(* IEC 61131-3 sources: daoli-st-library/DL_Motion (part 6) *)

(* ---- FB_DL_AxisCoggingFf.st ---- *)
(*==============================================================================
 * 组件名称 (Component)  : FB_DL_AxisCoggingFf
 * 所属子库 (Sublibrary) : DL_Motion
 * 当前版本 (Version)    : 1.0.0
 * 兼容性   (Platform)   : CODESYS 3.5+ / TwinCAT 3 / 汇川 InoProShop / 施耐德 Machine Expert
 *                         仅依赖 Standard.library（R_TRIG），零厂商私有库
 * 功能描述 (Function)   : 齿槽转矩前馈（按角度周期查表注入）。
 *                         把机械角等分成 72 个扇区（每扇区 5°），表内每格存该角度位置的补偿量；
 *                         运行时按当前角度取格、乘增益、限幅后以转矩前馈输出（% 额定）。
 *                         **学习与注入分离**（互斥锁存）：
 *                           注入态（bInjectEnable）：只读表 + 输出前馈，绝不改表；
 *                           学习态（bLearnEnable） ：只按"实测转矩指令"缓慢更新表内一格，绝不输出前馈；
 *                           两者同拍为真 → 锁存 eLearnConflict 并**两态全停**（既不改表也不输出），
 *                           避免"边学边补"形成正反馈自激。
 *                         三条固化纪律：
 *                           ① **相位取模防越界**：索引由角度除法取整后对 72 取模，负角再补 72，
 *                              结果恒落 0..71；角度非有限或超 ±1E6 度时当拍不判（防整数转换溢出）；
 *                           ② **注入限幅**：输出钳 ±fFfMaxPct，学习后的表格值同样钳在 ±fTableMaxPct；
 *                           ③ **学习率域闸**：fLearnRate 须在 (0, 1] 内，越域即锁存 eCfgIllegal
 *                              （大于 1 的学习率会使表格发散）。
 *                         验收向量：
 *                           ① 角度 0° → 索引 0；角度 5° → 索引 1；角度 355° → 索引 71
 *                           ② 角度 −5° → 索引 71（负角补模）
 *                           ③ 表[0] = 2.0 %、增益 1.0、限幅 5.0 → 前馈 2.0 %
 *                           ④ bInjectEnable 与 bLearnEnable 同拍为真 → eLearnConflict 锁存，输出 0
 * 接口     (Interface)  : 入 fAngleDeg 反馈机械角、bInjectEnable 注入使能、bLearnEnable 学习使能、
 *                         fTorqueRefPct 实测转矩（学习用观测值）、fFfGain 前馈增益、fFfMaxPct 注入限幅、
 *                         fTableMaxPct 表格值限幅、fLearnRate 学习率、bClear 清表沿、bReset 复位沿；
 *                         出 fFfOutPct 转矩前馈输出、iTableIdx 当前表索引（0..71）、bInjecting 注入中、
 *                         bLearning 学习中、bLearnConflict 学/注冲突锁存、bValid 输出有效、
 *                         eState 相、eCause 成因、bError 故障标志。
 * 边界     (Boundary)   : ① **属主边界（写死）：本件只做"角度周期前馈注入与表学习"，不输出位置/速度指令、
 *                         不参与轴使能与故障处理**——与 `FB_DL_AxisFrictionFf` 的分工：齿槽转矩是角度的
 *                         周期函数，摩擦转矩是速度的函数，两表互不替代（R47 边界声明）；
 *                         ② **状态枚举禁定义**：本件不引用任何轴状态枚举（R277），只消费角度引脚；
 *                         ③ **索引边界**：72 格字面量上界（R104），取模后恒在域内，另设显式钳位二次闸；
 *                         ④ **非有限闸**：角度/观测转矩非有限 → 当拍不判、不宣称（不锁存）；
 *                         ⑤ **锁存解除式**：bLearnConflict 与 eFault 仅由 bReset 上升沿解除（R228B），
 *                         bReset 为外部引脚、恒可达；
 *                         ⑥ 零全局耦合、零物理地址。
 * 分工声明 (Scope)      : 本件只管"齿槽转矩前馈"。不接管：摩擦前馈（属 FB_DL_AxisFrictionFf）、
 *                         反向间隙辨识（属 FB_DL_AxisBacklashIdent）、转矩环整定（属驱动侧）。
 * 来源标签 (Source Tag) : 自研线（与 AxisFrictionFf 成族）
 * 码表     (Codes)      : 本件不占用任何全局数字码位（零码位范式 R297）；诊断由 BOOL + ENUM 出口承担。
 * 红线自检 (Redline)    : R1 ✓ 零 GVL/VAR_EXTERNAL ｜ R2 ✓ 零 %I/%Q/%M ｜ R3 ✓ 纯 IEC 61131-3
 *                         R4 ✓ 取模 + 显式钳位 + 双限幅 + 学习率域闸 + 非有限闸 ｜ R5 ✓ 声明逐行同行双语注释
 *                         R6 ✓ ENUM+CASE 含 ELSE 兜底 ｜ R7 ✓ 两 R_TRIG 段 0 无条件刷新（本件无 TON）
 * 修订历史 (Revision)   : 2026-11-19  v1.0.0  R47 首版（批次 4 · 序号 20）
 *==============================================================================*)

TYPE E_DL_AcgState :
(
    eIdle  := 0,    // 待机相（两态皆关，输出 0） / Idle, both modes off, zero output
    eInject:= 10,   // 注入相（只读表输出前馈） / Injecting, table read only
    eLearn := 20,   // 学习相（只更新表，无输出） / Learning, table update only
    eFault := 90    // 故障相（等复位） / Fault, awaiting reset
);
END_TYPE

TYPE E_DL_AcgCause :
(
    eNone         := 0,   // 无异常 / No anomaly
    eCfgIllegal   := 1,   // 组态非法（学习率/限幅越域） / Illegal configuration
    eLearnConflict:= 2,   // 学习与注入同拍（锁存，两态全停） / Learn and inject together, latched
    eAngleBad     := 3,   // 角度非有限或超域（当拍不判） / Angle invalid, skipped this scan
    ePhaseBad     := 4    // 非法相位兜底 / Illegal phase fallback
);
END_TYPE

FUNCTION_BLOCK FB_DL_AxisCoggingFf
VAR_INPUT
    fAngleDeg    : LREAL := 0.0;      // 反馈机械角（可正可负） [°] / Feedback mechanical angle [°]
    bInjectEnable: BOOL := FALSE;     // 注入使能（只读表） [-] / Injection enable, table read only
    bLearnEnable : BOOL := FALSE;     // 学习使能（只改表） [-] / Learning enable, table write only
    fTorqueRefPct: LREAL := 0.0;      // 实测转矩（学习观测值） [% 额定] / Measured torque for learning [% rated]
    fFfGain      : LREAL := 1.0;      // 前馈增益，域 ≥ 0 [-] / Feed-forward gain, >= 0
    fFfMaxPct    : LREAL := 20.0;     // 注入限幅，域 > 0 [% 额定] / Injection clamp, > 0
    fTableMaxPct : LREAL := 30.0;     // 表格值限幅，域 > 0 [% 额定] / Table-value clamp, > 0
    fLearnRate   : LREAL := 0.01;     // 学习率，域 (0, 1] [-] / Learning rate, within (0, 1]
    bClear       : BOOL := FALSE;     // 清表沿（表格全置 0） [-] / Table-clear edge
    bReset       : BOOL := FALSE;     // 故障复位沿 [-] / Fault reset edge
END_VAR
VAR_OUTPUT
    fFfOutPct    : LREAL := 0.0;                          // 转矩前馈输出（已限幅） [% 额定] / Feed-forward output, clamped
    iTableIdx    : INT := 0;                              // 当前表索引（0..71） [-] / Present table index
    bInjecting   : BOOL := FALSE;                         // 注入中 [-] / Injecting
    bLearning    : BOOL := FALSE;                         // 学习中 [-] / Learning
    bLearnConflict : BOOL := FALSE;                       // 学/注冲突锁存（等复位） [-] / Learn-inject conflict, latched
    bValid       : BOOL := FALSE;                         // 输出有效（角度有效且注入态） [-] / Output valid
    eState       : E_DL_AcgState := E_DL_AcgState.eIdle;  // 相出口 [-] / Phase outlet
    eCause       : E_DL_AcgCause := E_DL_AcgCause.eNone;  // 成因出口（R190 归因唯一） [-] / Cause outlet
    bError       : BOOL := FALSE;                         // 故障标志（仅故障级成因） [-] / Error flag, fault level only
END_VAR
VAR
    _eState   : E_DL_AcgState := E_DL_AcgState.eIdle;    // 内部相（CASE 唯一写入目标） / Internal phase
    _eCause   : E_DL_AcgCause := E_DL_AcgCause.eNone;    // 成因锁存量 / Latched cause
    _bFault   : BOOL := FALSE;                           // 故障锁存位 / Latched fault bit
    _bConf    : BOOL := FALSE;                           // 学/注冲突锁存位 / Latched conflict bit
    _iIdx     : INT := 0;                                // 归一后的表索引（0..71） [-] / Normalised table index
    _iRaw     : INT := 0;                                // 取模前的索引 [-] / Index before normalisation
    _fOut     : LREAL := 0.0;                            // 输出工作值 [% 额定] / Output working value
    _fCell    : LREAL := 0.0;                            // 当格补偿量 [% 额定] / Cell compensation value
    _bAngOk   : BOOL := FALSE;                           // 角度有效性结论 / Angle validity result
    _bCfgBad  : BOOL := FALSE;                           // 组态非法当拍量 / Illegal configuration this scan
    _i        : INT := 0;                                // 清表循环下标 / Clear-loop index
    rtClear   : R_TRIG;                                  // 清表沿实例，段 0 无条件调用 / Clear edge instance
    rtReset   : R_TRIG;                                  // 复位沿实例，段 0 无条件调用 / Reset edge instance
    afTable   : ARRAY[0..71] OF LREAL;                   // 齿槽补偿表（72 格 = 5°/格，字面量上界） [% 额定] / Cogging table
END_VAR
VAR CONSTANT
    DL_ACG_NBINS   : INT := 72;          // 表格数（与数组字面量上界同源） [格] / Table bin count
    DL_ACG_BIN_DEG : LREAL := 5.0;       // 每格角度宽（360/72） [°] / Bin width in degrees
    DL_ACG_ANG_MAX : LREAL := 1000000.0; // 角度绝对值上限（防实数转整数溢出） [°] / Angle magnitude limit
    DL_ACG_EPS     : LREAL := 1.0E-12;   // 浮点判等容差 [-] / Equality tolerance
END_VAR

(* —— 段 0：组态闸 + 两沿无条件周期刷新（R228A；本件无 TON） —— *)
_bCfgBad := (fLearnRate <= 0.0) OR (fLearnRate > 1.0)                 // 学习率须在 (0, 1] / Learning rate within (0, 1]
         OR (fFfMaxPct <= 0.0) OR (fTableMaxPct <= 0.0)               // 两限幅须为正 / Both clamps positive
         OR (fFfGain < 0.0);                                          // 增益须非负 / Gain non-negative
rtClear(CLK := bClear);                                               // 清表沿 / Clear edge
rtReset(CLK := bReset);                                               // 复位沿 / Reset edge

(* —— 段 1：单拍/输出量预置（锁存量 _eCause/_bFault/_bConf/_iIdx 不入清单，R107） —— *)
fFfOutPct  := 0.0;                                                    // 前馈输出预置 / Feed-forward preset
bInjecting := FALSE;                                                  // 注入中预置 / Injecting preset
bLearning  := FALSE;                                                  // 学习中预置 / Learning preset
bValid     := FALSE;                                                  // 有效位预置 / Validity preset
bError     := FALSE;                                                  // 故障标志预清（R45 配对） / Error preset
_fOut      := 0.0;                                                    // 输出工作值预置 / Output working preset

(* —— 段 2：组态闸（非法即锁存） —— *)
IF _bCfgBad THEN
    _eCause := E_DL_AcgCause.eCfgIllegal;                             // 归因：组态非法 / Cause: illegal configuration
    _bFault := TRUE;                                                  // 锁存 / Latch
    _eState := E_DL_AcgState.eFault;                                  // 入故障相 / Enter fault phase
END_IF

(* —— 段 3：学/注冲突闸（同拍为真即锁存，两态全停） —— *)
IF bInjectEnable AND bLearnEnable THEN
    _bConf  := TRUE;                                                  // 冲突锁存 / Latch the conflict
    _bFault := TRUE;                                                  // 故障锁存 / Latch the fault
    _eCause := E_DL_AcgCause.eLearnConflict;                          // 归因：学/注冲突 / Cause: learn-inject conflict
    _eState := E_DL_AcgState.eFault;                                  // 入故障相 / Enter fault phase
END_IF

(* —— 段 4：迁出链与清表链（两条显式写出） —— *)
IF rtReset.Q THEN
    _bFault := FALSE;                                                 // 清故障锁存 / Clear fault latch
    _bConf  := FALSE;                                                 // 清冲突锁存 / Clear the conflict latch
    _eCause := E_DL_AcgCause.eNone;                                   // 清成因 / Clear cause
    _eState := E_DL_AcgState.eIdle;                                   // 回待机相 / Back to idle
END_IF
IF rtClear.Q THEN
    FOR _i := 0 TO 71 DO
        afTable[_i] := 0.0;                                           // 逐格清零（循环上界恒定） / Clear every bin
    END_FOR
END_IF

(* —— 段 5：索引归一（角度有限性 → 取整 → 取模 → 负角补模 → 显式钳位） —— *)
_bAngOk := NOT ((fAngleDeg <> fAngleDeg) OR ((fAngleDeg - fAngleDeg) <> (fAngleDeg - fAngleDeg)))
        AND (ABS(fAngleDeg) <= DL_ACG_ANG_MAX);                       // 有限且未超防溢出上限 / Finite and below the guard limit
IF _bAngOk THEN
    _iRaw := LREAL_TO_INT(TRUNC(fAngleDeg / DL_ACG_BIN_DEG));         // 取整到格号（截断向 0） / Truncate to a bin number
    _iIdx := _iRaw MOD DL_ACG_NBINS;                                  // 对格数取模 / Modulo the bin count
    IF _iIdx < 0 THEN
        _iIdx := _iIdx + DL_ACG_NBINS;                                // 负角补模（−5° → 71） / Negative angle wrapped
    END_IF
    IF _iIdx < 0 THEN
        _iIdx := 0;                                                   // 二次下钳（结构性冗余） / Second lower clamp
    ELSIF _iIdx > (DL_ACG_NBINS - 1) THEN
        _iIdx := DL_ACG_NBINS - 1;                                    // 二次上钳（结构性冗余） / Second upper clamp
    END_IF
    iTableIdx := _iIdx;                                               // 索引出口 / Index outlet
ELSE
    _eCause := E_DL_AcgCause.eAngleBad;                               // 归因：角度无效（当拍不判） / Cause: invalid angle
END_IF

(* —— 段 6：相迁移（注入 / 学习互斥；故障由段 4 迁出） —— *)
CASE _eState OF

E_DL_AcgState.eIdle:
    IF bInjectEnable AND (NOT bLearnEnable) THEN
        _eState := E_DL_AcgState.eInject;                              // 进注入相 / Enter injecting
    ELSIF bLearnEnable AND (NOT bInjectEnable) THEN
        _eState := E_DL_AcgState.eLearn;                               // 进学习相 / Enter learning
    END_IF

E_DL_AcgState.eInject:
    IF bLearnEnable THEN
        _eState := E_DL_AcgState.eIdle;                                // 学习被使能：先退注入（互斥由段 3 判冲突） / Leave injecting
    ELSIF NOT bInjectEnable THEN
        _eState := E_DL_AcgState.eIdle;                                // 失能：回待机 / Disabled, back to idle
    END_IF

E_DL_AcgState.eLearn:
    IF bInjectEnable THEN
        _eState := E_DL_AcgState.eIdle;                                // 注入被使能：先退学习 / Leave learning
    ELSIF NOT bLearnEnable THEN
        _eState := E_DL_AcgState.eIdle;                                // 失能：回待机 / Disabled, back to idle
    END_IF

E_DL_AcgState.eFault:
    ;                                                                  // 故障相：由段 4 复位沿迁出 / Exit via the reset edge

ELSE
    _eCause := E_DL_AcgCause.ePhaseBad;                                // 归因：非法相位 / Cause: illegal phase
    _bFault := TRUE;                                                   // 锁存 / Latch
    _eState := E_DL_AcgState.eFault;                                   // 强拉故障相 / Force fault phase

END_CASE

(* —— 段 7：注入（只读表；增益与限幅） —— *)
IF (_eState = E_DL_AcgState.eInject) AND _bAngOk THEN
    _fCell := afTable[_iIdx];                                           // 读当格补偿量 / Read the cell value
    _fOut  := _fCell * fFfGain;                                         // 乘增益 / Apply the gain
    IF _fOut > fFfMaxPct THEN
        _fOut := fFfMaxPct;                                             // 上限钳位 / Clamp high
    ELSIF _fOut < (0.0 - fFfMaxPct) THEN
        _fOut := 0.0 - fFfMaxPct;                                       // 下限钳位 / Clamp low
    END_IF
    bInjecting := TRUE;                                                 // 注入中 / Injecting
    bValid     := TRUE;                                                 // 输出有效 / Output valid
END_IF

(* —— 段 8：学习（只改表；观测转矩有限才更新；表值双限幅） —— *)
IF (_eState = E_DL_AcgState.eLearn) AND _bAngOk THEN
    IF NOT ((fTorqueRefPct <> fTorqueRefPct) OR ((fTorqueRefPct - fTorqueRefPct) <> (fTorqueRefPct - fTorqueRefPct))) THEN
        afTable[_iIdx] := afTable[_iIdx] + (fLearnRate * fTorqueRefPct);   // 梯度式更新（学习率已过域闸） / Gradient-style update
        IF afTable[_iIdx] > fTableMaxPct THEN
            afTable[_iIdx] := fTableMaxPct;                             // 表格上限钳位 / Table clamp high
        ELSIF afTable[_iIdx] < (0.0 - fTableMaxPct) THEN
            afTable[_iIdx] := 0.0 - fTableMaxPct;                       // 表格下限钳位 / Table clamp low
        END_IF
        bLearning := TRUE;                                              // 学习中 / Learning
    END_IF
END_IF

(* —— 段 9：出口单点映射（名实双出口，R191） —— *)
fFfOutPct      := _fOut;                                                // 前馈输出出口 / Feed-forward outlet
bLearnConflict := _bConf;                                               // 冲突锁存出口 / Conflict outlet
eState         := _eState;                                              // 相出口 / Phase outlet
eCause         := _eCause;                                              // 成因出口 / Cause outlet
bError         := _bFault;                                              // 故障标志 / Error flag

END_FUNCTION_BLOCK

(* ---- FB_DL_AxisDroopComp.st ---- *)
(*==============================================================================
 * 组件名称 (Component)  : FB_DL_AxisDroopComp
 * 所属子库 (Sublibrary) : DL_Motion
 * 当前版本 (Version)    : 1.0.0
 * 兼容性   (Platform)   : CODESYS 3.5 / TwinCAT 3 / 汇川 InoProShop / Machine Expert
 *                         仅依赖 Standard.library（R_TRIG），零厂商方言
 * 功能描述 (Function)   : 轴跟随误差前馈补偿：按速度段从补偿表取增益，折算位置前置量
 *                         fCompOut [mm] = 速度段增益 [mm per mm/s] × 速度给定 [mm/s]，
 *                         并钳在 ±fCompMax；用于抵消伺服刚度不足造成的跟随下垂。
 * 分工互引 (Boundary)   : FB_DL_AxisFollowErrGuard 是**保护件**（跟随误差超限即停），
 *                         本件是**补偿件**（前置量注入位置环，不产生任何停止动作）；
 *                         两者互不替代，禁把保护判据写进本件。
 *                         FB_DL_AxisFrictionFf 补偿摩擦力方向项，本件只补偿速度相关下垂。
 * 边界与语义披露 (Boundary disclosure) :
 *   1) 补偿表 8 段定长（DL_AC_SEG），段边界按 |fVelCmd| 等分 fVelSegMax，
 *      符号由速度给定方向携带（段内取绝对值查表，输出乘回方向），故负速也有补偿。
 *   2) 组态域闸（R151 全枚举）：fVelSegMax <= 0、fCompMax < 0、表内任一元素非有限或
 *      为负（负增益会让补偿反向加剧下垂）均判组态非法，锁存至复位沿 + 组态改对。
 *   3) 速度给定非有限属运行时信号失效：本拍不输出补偿（fCompOut := 0，安全侧不注入
 *      错误前置量），置信息级码，**不锁存**（不因一扫 NaN 让补偿永久失效）。
 *   4) 输出饱和（|补偿| 被 fCompMax 钳住）为信息级：饱和本身不改变补偿符号。
 * 故障码表 (Error codes) :
 *   16#0004_03F0 [故障级] 组态非法（段宽 / 补偿上限 / 表元素），补偿置 0
 *                 反证：补偿置 0 与「速度恰好为 0」输出组合相同，无码不可区分。
 *   16#0004_03F2 [信息级] 速度给定非有限，本拍不注入补偿（保持 0）
 *                 反证：补偿 0 与「低速段增益为 0」输出相同，需码位区分信号失效。
 *   16#0004_03F3 [信息级] 补偿量被上限钳位（bSaturated 同源可查）
 *                 反证：钳位后补偿与前一段恰好相同，无码不可观测。
 * 码位总账 (Code ledger) : 16#0004_03F0 用 ｜ 16#0004_03F2 / 03F3 用
 * 依赖     (Depends)    : 无 DL_ 内部依赖；Standard.library: R_TRIG
 * 红线自检 (Redline)    : R1 ✓ 零全局变量 ｜ R2 ✓ 零 %I/%Q ｜ R3 ✓ 纯 IEC 61131-3
 *                         R4 ✓ 段索引钳位无越界 / 非有限三判 / 除子由域闸保证 > 0
 *                         R5 ✓ 全变量双语同行注释 ｜ R6 ✓ 三态 ENUM + ELSE 兜底
 *                         R7 ✓ 一沿实例主体最前部无条件刷新
 * 修订历史 (Revision)   : 2026-11-22  v1.0.0  首版入库（R69 构建轮 · 批 3 · N8）
 *============================================================================*)

(*-----------------------------------------------------------------------------
 * 枚举: E_DL_DroopState（归属 DL_Motion，与 FB_DL_AxisDroopComp 同文件）
 *----------------------------------------------------------------------------*)
TYPE E_DL_DroopState :
(
    eOff   := 0,      // 未使能：补偿恒 0 / Disabled, compensation is zero
    eRun   := 10,     // 补偿中：按速度段查表 / Compensating by speed segment
    eFault := 99      // 组态锁存：补偿恒 0 / Config latched, compensation forced to zero
);
END_TYPE

(*==============================================================================
 * 功能块: FB_DL_AxisDroopComp
 * 调用约定: 每个扫描周期无条件调用一次。
 *============================================================================*)
FUNCTION_BLOCK FB_DL_AxisDroopComp
VAR_INPUT
    fVelCmd    : REAL;                          // 速度给定 [mm/s] / velocity setpoint [mm/s]
    afSegGain  : ARRAY[0..7] OF REAL;           // 8 段补偿增益 [mm per mm/s]，必须 >= 0 / per-segment droop gain
    fVelSegMax : REAL := 1000.0;                // 补偿表覆盖的最高速度 [mm/s]，<= 0 组态非法 / table velocity span
    fCompMax   : REAL := 2.0;                   // 补偿量上限 [mm]，< 0 组态非法 / compensation magnitude ceiling [mm]
    bEnable    : BOOL := TRUE;                  // 使能 / enable
    bReset     : BOOL;                          // 上升沿：清组态锁存 / rising edge clears the config latch
END_VAR
VAR_OUTPUT
    fCompOut   : REAL;                          // 位置前置补偿量 [mm]（含速度方向符号）/ position feed-forward [mm]
    nSegIdx    : INT;                           // 命中补偿段号 [段]，0..7 / hit segment index
    bSaturated : BOOL;                          // 补偿量被上限钳位 / compensation clamped at the ceiling
    bVelValid  : BOOL;                          // 本拍速度给定有限 / velocity setpoint finite this scan
    bError     : BOOL;                          // 故障标志（组态锁存）/ fault flag
    uErrorId   : UDINT;                         // 故障码，0 = 无故障 / error code, 0 = none
    eState     : E_DL_DroopState;               // 当前状态（供 HMI 诊断）/ current state
END_VAR
VAR
    fbTrigReset : R_TRIG;                       // 复位沿检测实例 / reset edge detector
    eStateInt   : E_DL_DroopState;              // 主状态机内部当前态 / internal state
    fVelAbs     : REAL;                         // 速度绝对值 [mm/s]（查表用）/ absolute velocity for the lookup
    fSegSpan    : REAL;                         // 单段速度宽度 [mm/s]（除子，域闸保证 > 0）/ segment width, the divisor
    fGainEff    : REAL;                         // 命中段增益 [mm per mm/s] / hit segment gain
    fCompRaw    : REAL;                         // 未钳补偿量 [mm] / unclamped compensation
    nIdx        : INT;                          // 表遍历游标 [段] / table cursor
    bVelBad     : BOOL;                         // 速度给定非有限 / velocity non-finite
    bCfgBad     : BOOL;                         // 本拍组态非法 / config illegal this scan
    bCfgLatch   : BOOL;                         // 组态锁存（复位沿 + 组态改对解除）/ config latch
    bErrorInt   : BOOL;                         // 本拍故障置位累加 / fault set accumulator
    bFirstScan  : BOOL := TRUE;                 // 上电首扫标志 / first-scan flag
END_VAR
VAR CONSTANT
    DL_AC_SEG     : INT := 8;                   // 补偿表段数 [段]，与数组维度一致 / segment count
    DL_AC_FIN_LIM : REAL := 1.0E30;             // REAL 幅值兜底判界 / REAL magnitude bound
    DL_AC_NEG_EPS : REAL := 0.0;                // 增益负值判界（0 为合法端点）/ gain negativity bound, zero is legal
END_VAR

(*------------------------------------------------------------------------------
 * 段 1｜无条件刷新区（红线 R7）：一沿实例位于主体最前部
 *      Unconditional refresh: the edge instance at the very top
 *-----------------------------------------------------------------------------*)
fbTrigReset(CLK := bReset);

(* 段 2｜上电首扫：状态与输出落安全侧 / first-scan init *)
IF bFirstScan THEN
    eStateInt  := E_DL_DroopState.eOff;
    fCompOut   := 0.0;
    bFirstScan := FALSE;
END_IF

(* 段 3｜每拍预清（FB32-1）：单拍标志与派生量 / per-scan preset *)
bErrorInt  := FALSE;
bSaturated := FALSE;

(*------------------------------------------------------------------------------
 * 段 4｜组态域闸（R151 全枚举）：段宽 / 上限 / 表内 8 个元素逐一非有限与负值判
 *      Config gate over the span, the ceiling and every table element
 *      解除路径（R152 自证可达）：复位沿 AND 组态非法条件全部消失
 *-----------------------------------------------------------------------------*)
bCfgBad := (fVelSegMax <= 0.0) OR (fVelSegMax <> fVelSegMax)
           OR (fCompMax < 0.0) OR (fCompMax <> fCompMax);
FOR nIdx := 0 TO (DL_AC_SEG - 1) DO
    IF (afSegGain[nIdx] <> afSegGain[nIdx])
       OR ((afSegGain[nIdx] - afSegGain[nIdx]) <> (afSegGain[nIdx] - afSegGain[nIdx]))
       OR (ABS(afSegGain[nIdx]) >= DL_AC_FIN_LIM)
       OR (afSegGain[nIdx] < DL_AC_NEG_EPS) THEN
        bCfgBad := TRUE;                        // 表元素非法：任一项即整表不可信 / any bad element invalidates the table
    END_IF
END_FOR

IF bCfgBad THEN
    bCfgLatch := TRUE;
END_IF
IF fbTrigReset.Q AND (NOT bCfgBad) THEN
    bCfgLatch := FALSE;                         // 组态锁存解除 / config latch cleared
    uErrorId  := 16#0000_0000;                  // 码位随解除归零 / code cleared with the latch
END_IF
IF bCfgLatch THEN
    uErrorId  := 16#0004_03F0;                  // 故障级：组态非法 / fault: illegal configuration
    bErrorInt := TRUE;                          // R45 配对 / paired with the code
    eStateInt := E_DL_DroopState.eFault;
END_IF

(*------------------------------------------------------------------------------
 * 段 5｜主状态机（红线 R6）：ENUM + CASE + ELSE 兜底
 *-----------------------------------------------------------------------------*)
CASE eStateInt OF

    E_DL_DroopState.eOff:
        IF bEnable AND (NOT bCfgLatch) THEN
            eStateInt := E_DL_DroopState.eRun;
        END_IF

    E_DL_DroopState.eRun:
        IF (NOT bEnable) OR bCfgLatch THEN
            eStateInt := E_DL_DroopState.eOff;
        END_IF

    E_DL_DroopState.eFault:
        IF fbTrigReset.Q AND (NOT bCfgBad) THEN
            bCfgLatch := FALSE;
            uErrorId  := 16#0000_0000;
            eStateInt := E_DL_DroopState.eOff;
        END_IF

    ELSE
        (* 非法状态拦截 / illegal state interception *)
        eStateInt := E_DL_DroopState.eFault;
        uErrorId  := 16#0004_03F0;
        bErrorInt := TRUE;

END_CASE;

(*------------------------------------------------------------------------------
 * 段 6｜速度段查表与补偿折算
 *      Segment lookup and the compensation folding
 *-----------------------------------------------------------------------------*)
bVelBad  := (fVelCmd <> fVelCmd)
            OR ((fVelCmd - fVelCmd) <> (fVelCmd - fVelCmd))
            OR (ABS(fVelCmd) >= DL_AC_FIN_LIM);
bVelValid := (NOT bVelBad) AND (NOT bCfgLatch);
fCompOut  := 0.0;                               // 缺省不注入（安全侧）/ default no injection
nSegIdx   := 0;
fGainEff  := 0.0;

IF bVelValid AND bEnable AND (eStateInt = E_DL_DroopState.eRun) THEN
    IF fVelCmd >= 0.0 THEN
        fVelAbs := fVelCmd;                     // 正方向 [mm/s] / positive direction
    ELSE
        fVelAbs := -fVelCmd;                    // 取绝对值查表（符号在出口乘回）[mm/s] / absolute value for the lookup
    END_IF
    fSegSpan := fVelSegMax / INT_TO_REAL(DL_AC_SEG);                 // 单段宽（除子为常数 8 > 0）[mm/s] / segment width
    IF fVelAbs > fVelSegMax THEN
        fVelAbs := fVelSegMax;                  // 实数域先钳制再转整型（R151 防方向翻转）/ clamp in the real domain before the cast
    END_IF
    nSegIdx  := REAL_TO_INT(fVelAbs / fSegSpan);                     // 段号（除子 > 0 且已钳制）/ segment index after clamping
    IF nSegIdx >= DL_AC_SEG THEN
        nSegIdx := DL_AC_SEG - 1;               // 超表按末段钳位（禁越界访问）/ clamp to the last segment
    ELSIF nSegIdx < 0 THEN
        nSegIdx := 0;                           // 负段号防御，结构性不可达 / negative guard, unreachable
    END_IF
    fGainEff := afSegGain[nSegIdx];             // 命中段增益 [mm per mm/s] / hit gain
    fCompRaw := fGainEff * fVelCmd;             // 未钳补偿（含方向符号）[mm] / raw compensation with direction
    IF fCompRaw > fCompMax THEN
        fCompOut   := fCompMax;                 // 正向饱和 [mm] / saturated high
        bSaturated := TRUE;
        uErrorId   := 16#0004_03F3;             // 信息级：补偿被钳位 / info: compensation clamped
    ELSIF fCompRaw < -fCompMax THEN
        fCompOut   := -fCompMax;                // 负向饱和 [mm] / saturated low
        bSaturated := TRUE;
        uErrorId   := 16#0004_03F3;             // 信息级：补偿被钳位 / info: compensation clamped
    ELSE
        fCompOut   := fCompRaw;                 // 域内直通 [mm] / in-domain pass-through
    END_IF
ELSIF bVelBad THEN
    uErrorId := 16#0004_03F2;                   // 信息级：速度非有限，不注入（不锁存）/ info: non-finite velocity
END_IF

(*------------------------------------------------------------------------------
 * 段 7｜输出单一出口（范式 P-05）
 *      Single output exit
 *-----------------------------------------------------------------------------*)
bError := bErrorInt OR bCfgLatch;
eState := eStateInt;
END_FUNCTION_BLOCK

(* ---- FB_DL_AxisDualFeedbackGuard.st ---- *)
(*==============================================================================
 * 组件名称 (Component)  : FB_DL_AxisDualFeedbackGuard
 * 所属子库 (Sublibrary) : DL_Motion
 * 当前版本 (Version)    : 1.0.0
 * 兼容性   (Platform)   : CODESYS 3.5+ / TwinCAT 3 / 汇川 InoProShop / 施耐德 Machine Expert
 *                         仅依赖 Standard.library（TON / R_TRIG / ABS），零厂商私有库
 * 功能描述 (Function)   : 单轴双反馈交叉校核。把电机侧位置 fPosMotor 与负载侧位置 fPosLoad
 *                         各自乘标定系数换算到同一工程单位后求偏差 fDev，并按幅值与持续时间
 *                         分级：|fDev| 超 fDevWarn → 维护级预警（bWarn）；超 fDevAlarm 且持续
 *                         tDevConfirm → 故障锁存。另做极性装反识别：偏差方向与参考运动方向
 *                         同号、且偏差每拍增量超 fSlopeThr 时归因 ePolarity（区别于打滑——
 *                         打滑时偏差随运动累积但方向与运动一致而增量平稳，装反时增量陡增）。
 * 接口     (Interface)  : 输入 fPosMotor 电机侧位置、fPosLoad 负载侧位置、fScaleMotor / fScaleLoad
 *                         两侧标定系数、fDevWarn 预警阈值、fDevAlarm 故障阈值、tDevConfirm 故障
 *                         确认时间、fSlopeThr 偏差每拍增量阈值、fVelRefMms 参考运动速度（方向
 *                         判据）、bReset 复位；输出 fDev 换算后偏差、bWarn 维护级预警、bGuardOk
 *                         校核通过、eState / eCause / bError / nErrId。
 * 边界     (Boundary)   : ① 组态闸：fScaleMotor / fScaleLoad 的绝对值 <= DL_FLOAT_EPS（防零增益
 *                         静默把偏差算成 0）、fDevWarn <= 0.0、fDevAlarm <= fDevWarn、
 *                         tDevConfirm <= T#0S、fSlopeThr < 0.0 或任一浮点引脚 NaN → 故障锁存；
 *                         ② **本件不定义轴状态枚举、不发运动指令**（轴状态唯一属主 `I_DL_MotionAxis`），
 *                         只读位置与速度参考，只输出校核结论；
 *                         ③ 偏差每拍增量以「每拍工程单位增量」为单位：任务周期固定时它与斜率
 *                         成正比，fSlopeThr 按该口径标定（比值约定见头注释遗留假设）；
 *                         ④ TON 两枚（预警/故障确认）+ R_TRIG 一枚段 0 无条件周期刷新；
 *                         ⑤ 故障相迁出唯一路径 = bReset 上升沿；⑥ 零全局耦合（无 GVL / 无物理地址）。
 * 分工声明 (Scope)      : 与 `FB_DL_GantrySyncAxis`（双**轴**同步偏差）分工 —— 本件是**单轴双反馈**
 *                         （电机侧 vs 负载侧），判「同一根轴的两把尺是否一致」；那件判「两根轴的
 *                         位置是否同步」。二者输入维度不同，禁止互相替代。
 * 遗留假设 (Assumption) : 【R95 三句声明】① 代理值 = 偏差每拍增量（未引入任务周期引脚）；
 *                         ② 覆盖范围 = 任务周期 1 ms ~ 20 ms 的常规运动任务；③ 覆盖不到的区间
 *                         （< 1 ms 的高速插补任务）由调用方负责：此时每拍增量被任务周期压缩，
 *                         fSlopeThr 需由调用方按周期比例放大，否则极性识别灵敏度下降。
 * 解除式   (Release)    : bReset 上升沿 ∧ 组态合法 ∧ |fDev| < fDevWarn（当拍量，R240 范式）。
 *                         自证可满足（终审两式 1）：解除式只含当拍偏差比较与组态闸，两枚 TON
 *                         的 IN 由当拍阈值判据派生，偏差回落即 Q 落假，无恒假因子。
 * 码表     (Codes)      : 16#0004_03B4 故障级：双反馈校核故障总码（组态非法 / 偏差超限确认 /
 *                         极性装反 / 非法相位），锁存至 bReset 上升沿，归因由 eCause 承载；
 *                         16#0004_04B4 信息级：维护级预警（|fDev| 超 fDevWarn 但未达故障）。
 *                         加码反证（R90）：预警相 fDev 仍为小值、bError 为假，若只靠 bWarn 布尔
 *                         位则该退化不进报警台账（HMI 只归档带码事件），故立一码。
 *                         码段说明：0004 段故障子带 03xx / 信息子带 04xx，本件取 03B4 / 04B4
 *                         （源码实扫该两槽为空，续接同子带已用最大值，未回填碎片孔洞）。
 * 开源溯源 (Origin)     : 道莅自研 clean-room（参考双反馈交叉校核与极性判别参数域，零代码行复制；
 *                         t1-6-plcopen 族）
 * 修订历史 (Revision)   : 2026-11-19  v1.0.0  R45 首版（批次 2 · 序号 10）
 *==============================================================================*)

TYPE E_DL_DfgState :
(
    eIdle  := 0,     // 未取得有效反馈，等待首拍 / Idle, awaiting first valid feedback
    eRun   := 10,    // 校核运行 / Guard running
    eFault := 90     // 故障锁存相 / Fault latched phase
);
END_TYPE

TYPE E_DL_DfgCause :
(
    eNone       := 0,   // 无故障成因 / No cause
    eCfgIllegal := 1,   // 组态非法 / Illegal configuration
    eDevLimit   := 2,   // 偏差超故障阈值且确认时间到 / Deviation over alarm limit confirmed
    ePolarity   := 3,   // 极性装反（偏差随运动同号且增量陡增） / Polarity reversed
    ePhaseBad   := 4    // 非法相位兜底 / Illegal phase fallback
);
END_TYPE

FUNCTION_BLOCK FB_DL_AxisDualFeedbackGuard
VAR_INPUT
    fPosMotor   : REAL := 0.0;          // 电机侧位置（编码器计数或已换算值） [cnt] / Motor-side position in encoder counts [cnt]
    fPosLoad    : REAL := 0.0;          // 负载侧位置（光栅尺或第二编码器） [mm] / Load-side position from scale [mm]
    fScaleMotor : REAL := 0.001;        // 电机侧标定系数，绝对值须 > DL_FLOAT_EPS [mm/cnt] / Motor-side scale, |value| > epsilon [mm/cnt]
    fScaleLoad  : REAL := 1.0;          // 负载侧标定系数，绝对值须 > DL_FLOAT_EPS [mm/mm] / Load-side scale, |value| > epsilon [mm/mm]
    fDevWarn    : REAL := 0.05;         // 维护级预警阈值，域 > 0.0 [mm] / Maintenance warning threshold, domain > 0.0 [mm]
    fDevAlarm   : REAL := 0.20;         // 故障阈值，域 > fDevWarn [mm] / Fault threshold, domain > fDevWarn [mm]
    tDevConfirm : TIME := T#200MS;      // 故障确认时间，域 > T#0S [ms] / Fault confirm time, domain > T#0S [ms]
    fSlopeThr   : REAL := 0.02;         // 偏差每拍增量阈值（极性判据），域 >= 0.0 [mm/拍] / Deviation increment per scan threshold [mm/scan]
    fVelRefMms  : REAL := 0.0;          // 参考运动速度（仅用符号判方向） [mm/s] / Reference velocity, sign used for direction [mm/s]
    bReset      : BOOL := FALSE;        // 复位命令，上升沿清故障 [-] / Reset command, rising edge clears fault
END_VAR
VAR_OUTPUT
    fDev        : REAL;                 // 换算到同一单位后的偏差（电机侧 − 负载侧） [mm] / Deviation after unit conversion [mm]
    bWarn       : BOOL;                 // 维护级预警（未达故障） [-] / Maintenance warning, below fault level
    bGuardOk    : BOOL;                // 校核通过（偏差在预警带内且无故障） [-] / Guard passed
    eState      : E_DL_DfgState;        // 状态出口，段 6 单点映射 / State outlet
    eCause      : E_DL_DfgCause;        // 故障成因出口（R190 归因唯一） / Fault cause outlet
    bError      : BOOL;                 // 故障锁存标志 [-] / Fault latch flag
    nErrId      : UDINT;               // 事件码，0 = 无事件 / Event code, 0 = no event
END_VAR
VAR
    _eState     : E_DL_DfgState := E_DL_DfgState.eIdle;    // 内部相位（CASE 唯一写入目标） / Internal phase
    _eCause     : E_DL_DfgCause := E_DL_DfgCause.eNone;    // 故障成因锁存（锁存量） / Latched cause
    tonWarn     : TON;                  // 预警确认计时，段 0 无条件调用 / Warning timer
    tonAlarm    : TON;                  // 故障确认计时，段 0 无条件调用 / Alarm confirm timer
    rtReset     : R_TRIG;               // 复位沿实例，段 0 无条件调用 / Reset edge
    _fMotorMm   : REAL;                 // 电机侧换算位置 [mm] / Motor-side position in millimetres
    _fLoadMm    : REAL;                 // 负载侧换算位置 [mm] / Load-side position in millimetres
    _fDevPrev   : REAL;                 // 上拍偏差快照（锁存量） [mm] / Previous-scan deviation snapshot
    _fDevStep   : REAL;                 // 本拍偏差增量 [mm] / Deviation increment this scan
    _fDev       : REAL;                 // 本拍换算偏差中间量（段 0 派生，段 8 映射到输出） [mm] / Deviation intermediate, derived in seg 0, mapped to output in seg 8
    _bPolSame   : BOOL;                 // 偏差符号与运动方向同号当拍量 [-] / Deviation sign matches motion sign
    _bPolSteep  : BOOL;                 // 偏差增量超阈值当拍量 [-] / Deviation increment above threshold
    _bNonFin    : BOOL;                 // 输入非有限当拍量 [-] / Non-finite input this scan
    _bCfgBad    : BOOL;                 // 组态非法当拍量 [-] / Illegal configuration
    _bFault     : BOOL;                 // 故障锁存位（锁存量） / Latched fault bit
    _uFault     : UDINT;                // 故障码锁存（锁存量） / Latched fault code
    _uInfo      : UDINT;                // 信息码，每拍重算 / Info code, recomputed each scan
END_VAR
VAR CONSTANT
    DL_FLOAT_EPS : REAL := 1.0E-6;      // 浮点判零容差（标定系数与判据统一口径） [无量纲] / Float epsilon for zero tests
END_VAR

(* —— 段 0：当拍量派生 + 定时器与沿实例无条件周期刷新 —— *)
_fMotorMm := fPosMotor * fScaleMotor;                                    // 电机侧换算到 mm / Motor side converted to millimetres
_fLoadMm  := fPosLoad * fScaleLoad;                                      // 负载侧换算到 mm / Load side converted to millimetres
_fDev     := _fMotorMm - _fLoadMm;                                       // 偏差 = 电机侧 − 负载侧 [mm] / Deviation, motor minus load
_fDevStep := _fDev - _fDevPrev;                                          // 本拍偏差增量 [mm/拍] / Deviation increment per scan
_bNonFin  := (fPosMotor <> fPosMotor) OR (fPosLoad <> fPosLoad)          // NaN 自反判（判等禁令唯一例外） / NaN self-reflexive tests
          OR (fScaleMotor <> fScaleMotor) OR (fScaleLoad <> fScaleLoad)  // 标定系数 NaN 判 / Scale NaN tests
          OR (fVelRefMms <> fVelRefMms) OR (fSlopeThr <> fSlopeThr);     // 方向与阈值 NaN 判 / Direction and threshold NaN tests
_bCfgBad  := (ABS(fScaleMotor) <= DL_FLOAT_EPS) OR (ABS(fScaleLoad) <= DL_FLOAT_EPS)   // 零增益闸（R151 覆盖每个参与引脚） / Zero-gain gate
             OR (fDevWarn <= 0.0) OR (fDevAlarm <= fDevWarn)                           // 阈值几何闸 / Threshold geometry gate
             OR (tDevConfirm <= T#0S) OR (fSlopeThr < 0.0);                            // 时间与增量阈值闸 / Time and increment gates
_bPolSame := ((_fDev > 0.0) AND (fVelRefMms > 0.0)) OR ((_fDev < 0.0) AND (fVelRefMms < 0.0));   // 偏差与运动同号 / Deviation sign equals motion sign
_bPolSteep := ABS(_fDevStep) > fSlopeThr;                                                      // 增量陡增判据 / Steep increment criterion
rtReset(CLK := bReset);                                                                        // 复位沿，每拍必调（R228A） / Reset edge
tonWarn(IN := ABS(_fDev) > fDevWarn, PT := tDevConfirm);                                       // 预警确认计时（IN 由判据派生） / Warning timer
tonAlarm(IN := ABS(_fDev) > fDevAlarm, PT := tDevConfirm);                                     // 故障确认计时 / Alarm confirm timer

(* —— 段 1：单拍量预清零（锁存量与快照量不入清单，R107） —— *)
_uInfo    := 16#0000_0000;         // 信息码每拍重算 / Info recomputed every scan
bWarn     := FALSE;                // 预警位每拍预清 / Warning preset
bGuardOk  := FALSE;                // 通过位每拍预清 / Pass flag preset
nErrId    := 16#0000_0000;         // 事件码缺省无事件 / Event code default none
bError    := FALSE;                // 故障标志每拍预清，故障分支同拍置位（R45 配对） / Flag preset

(* —— 段 2：复位沿 + 组态域闸 + 非有限闸 —— *)
IF rtReset.Q THEN                                                        // 当拍复位沿 / current-scan reset edge
    _bFault := FALSE;                                                    // 清故障锁存位（锁存量） / Clear fault latch
    _uFault := 16#0000_0000;                                             // 清故障锁存码（锁存量） / Clear latched code
    _eCause := E_DL_DfgCause.eNone;                                      // 清成因（锁存量） / Clear latched cause
    IF _eState = E_DL_DfgState.eFault THEN
        _eState := E_DL_DfgState.eIdle;                                  // 故障相迁出唯一路径 / Sole exit from fault phase
    END_IF
END_IF
IF _bCfgBad THEN                                                         // 组态域闸 / Configuration gate
    _uFault := 16#0004_03B4;                                             // 故障级：双反馈校核故障总码 / Fault-level: guard fault code
    _bFault := TRUE;
    bError  := TRUE;                                                     // 故障标志同拍置位（R45 配对） / Error flag set same scan
    _eCause := E_DL_DfgCause.eCfgIllegal;                                // 归因：组态非法 / Cause: illegal configuration
END_IF
IF (NOT _bFault) AND _bNonFin THEN                                       // 输入非有限 / Non-finite input
    _uFault := 16#0004_03B4;
    _bFault := TRUE;
    bError  := TRUE;
    _eCause := E_DL_DfgCause.eDevLimit;                                  // 归因：偏差不可信（非有限并入超限） / Cause: deviation untrustworthy, folded into limit
END_IF

(* —— 段 3：极性装反识别（先于幅值分级判，避免装反被误归因为打滑） —— *)
IF (NOT _bFault) AND _bPolSame AND _bPolSteep AND (ABS(_fDev) > fDevWarn) THEN
    _uFault := 16#0004_03B4;
    _bFault := TRUE;
    bError  := TRUE;
    _eCause := E_DL_DfgCause.ePolarity;                                  // 归因：极性装反 / Cause: polarity reversed
END_IF

(* —— 段 4：幅值分级（预警=维护级信息；故障=确认窗到） —— *)
IF (NOT _bFault) THEN
    IF tonAlarm.Q THEN                                                   // 超故障阈值且确认窗到 / Over alarm limit confirmed
        _uFault := 16#0004_03B4;
        _bFault := TRUE;
        bError  := TRUE;
        _eCause := E_DL_DfgCause.eDevLimit;                              // 归因：偏差超限 / Cause: deviation over limit
    ELSIF ABS(_fDev) > fDevWarn THEN                                     // 预警带（维护级，不锁故障） / Warning band, maintenance level
        bWarn := TRUE;                                                   // 预警位 / Warning flag
        _uInfo := 16#0004_04B4;                                          // 信息级：维护级预警 / Info: maintenance warning
    ELSE
        bGuardOk := TRUE;                                                // 预警带内：校核通过 / Inside band, guard passed
    END_IF
END_IF

(* —— 段 5：偏差快照更新（主体末行，跨拍纪律） —— *)
_fDevPrev := _fDev;                                                      // 偏差快照（本拍末更新） / Deviation snapshot at body end

(* —— 段 6：故障解除式（R240 全当拍量） —— *)
IF rtReset.Q AND (NOT _bCfgBad) AND (ABS(_fDev) < fDevWarn) THEN
    _bFault := FALSE;                                                    // 清故障锁存位（锁存量） / Clear fault latch
    _uFault := 16#0000_0000;                                             // 清故障锁存码（锁存量） / Clear latched code
    _eCause := E_DL_DfgCause.eNone;                                      // 清成因（锁存量） / Clear latched cause
END_IF

(* —— 段 6A：故障锁存相位迁移闸 —— *)
IF _bFault AND (_eState <> E_DL_DfgState.eFault) THEN
    _eState := E_DL_DfgState.eFault;                                     // 锁存即入故障相 / Latch enters fault phase
END_IF

(* —— 段 7：相位机（ENUM 全成员显式标签 + ELSE 兜底，R128） —— *)
CASE _eState OF

E_DL_DfgState.eIdle:
    IF (NOT _bNonFin) AND (NOT _bCfgBad) AND (rtReset.Q OR bGuardOk OR bWarn) THEN   // 出口 1：偏差可算且已判定（复位后首拍或已出结论） / Deviation computable and judged
        _eState := E_DL_DfgState.eRun;
    ELSIF _bFault THEN                                                   // 出口 2：故障锁存 / Fault latched
        _eState := E_DL_DfgState.eFault;
    END_IF

E_DL_DfgState.eRun:
    IF rtReset.Q AND (NOT _bFault) THEN                                  // 出口 1：运行相收到复位沿 → 回观测相重采样一次 / Reset re-arms the guard
        _eState := E_DL_DfgState.eIdle;
    ELSIF _bFault THEN                                                   // 出口 2：故障锁存 / Fault latched
        _eState := E_DL_DfgState.eFault;
    END_IF

E_DL_DfgState.eFault:
    ;                                                                     // 故障相：仅段 6 复位沿可迁出 / Only the reset edge leaves this phase

ELSE
    _uFault := 16#0004_03B4;                                             // 故障级：非法相位兜底（归并总码） / Illegal-phase fallback
    _bFault := TRUE;
    bError  := TRUE;
    _eCause := E_DL_DfgCause.ePhaseBad;                                  // 归因：非法相位 / Cause: illegal phase
    _eState := E_DL_DfgState.eFault;

END_CASE

(* —— 段 8：出口单点映射（名实同源；锁存码回放；故障相安全侧） —— *)
IF _bFault THEN
    bWarn    := FALSE;                                                   // 故障相不再宣称「仅预警」 / No warning claim in fault
    bGuardOk := FALSE;                                                   // 故障相校核不通过 / Guard failed in fault
END_IF
IF _bFault THEN
    nErrId := _uFault;                                                   // 故障锁存码回放 / Replay latched fault code
ELSE
    nErrId := _uInfo;                                                    // 信息码 / Info code
END_IF
bError := _bFault;                                                       // 故障标志与锁存同源（名实双出口，R191） / Flag from latch
fDev    := _fDev;                                                               // 偏差输出每拍赋值（名实同源） / Deviation output assigned every scan
eState := _eState;                                                       // 状态出口 / State outlet
eCause := _eCause;                                                       // 成因出口 / Cause outlet

END_FUNCTION_BLOCK

(* ---- FB_DL_AxisEncoderPulseLostScore.st ---- *)
(*==============================================================================
 * 组件名称 (Component)  : FB_DL_AxisEncoderPulseLostScore
 * 所属子库 (Sublibrary) : DL_Motion
 * 当前版本 (Version)    : 1.0.0
 * 兼容性   (Platform)   : CODESYS 3.5+ / TwinCAT 3 / 汇川 InoProShop / 施耐德 Machine Expert
 *                         仅依赖 Standard.library（R_TRIG / ABS / MIN / MAX），零厂商私有库
 * 功能描述 (Function)   : 编码器脉冲丢失率在线评分分档。调用方在观测窗内累计脉冲数
 *                         nPulseCntWindow（窗口起点清零，由调用方负责）与本窗期望脉冲数
 *                         fExpectWindow（= |参考速度| × 每毫米脉冲数 × 窗口时长，由调用方换算）。
 *                         本件在 bWindowEnd 上升沿取一次快照，算比值 fRatio = 实测/期望，
 *                         再折成 0~100 分：fRatio >= 1.0 记 100 分；fRatio 在 [0,1) 段线性
 *                         衰减到 0 分（100 × fRatio）；fRatio > 1.0 按 100 分封顶（超发不奖分，
 *                         但另出 bOverRun 提示，防"丢脉冲与多脉冲相互掩盖"）。
 *                         评分分三档：>= nScoreGood 良好、>= nScoreWarn 关注、< nScoreWarn 劣化。
 * 接口     (Interface)  : 输入 nPulseCntWindow 窗内实测脉冲数、fExpectWindow 窗内期望脉冲数、
 *                         bWindowEnd 窗口结束沿、fRatioMin 有效比值下界（防期望值过小病态放大）、
 *                         nScoreGood / nScoreWarn 分档线；输出 fRatio 实测/期望、nScore 0~100、
 *                         eGrade 分档、bValid 本窗评分有效、eState / bError。
 * 边界     (Boundary)   : ① **属主边界（写死）：本件只评分，不判故障、不发报警、不改轴**。
 *                         故障级判定唯一属主为轴级监控链（`FB_DL_AxisFollowingErrorMonitor` 等）；
 *                         本件输出 nScore / eGrade 供上层做趋势与维护决策。
 *                         ② 组态闸：nScoreGood <= nScoreWarn、分档线 > 100 或 < 0、
 *                         fRatioMin <= 0.0、fExpectWindow 为 NaN → 故障（ELSE 兜底 + 成因归因）。
 *                         ③ 期望值为 0 或低于 fExpectWindow 下界 → 本窗不评分（bValid=FALSE，
 *                         nScore 保持上窗值不清零），并在 eCause 说明"激励不足"，严禁把
 *                         "无期望"记成 100 分（那会把停机的轴伪装成健康）。
 *                         ④ R_TRIG 一枚段 0 无条件周期刷新；无 TON，故无跨相不复位风险。
 *                         ⑤ 零全局耦合（无 GVL / 无 VAR_EXTERNAL / 无物理地址）。
 * 分工声明 (Scope)      : 与 `FB_DL_FrequencyMeasure`（测频）分工——那件给频率本身，本件给
 *                         "窗内实测/期望"的**比率与评分**，输入是已由调用方累计的脉冲计数。
 * 来源标签 (Source Tag) : T1-6 ◐（开源参考：脉冲丢失率在线评估参数域，零代码行复制）
 * 解除式   (Release)    : 本件无锁存故障相：bError 每拍重算（组态非法/非有限即置），
 *                         组态修正后下一拍自动消失——信息级与故障级的边界写死在此（R189 例外条款：
 *                         无锁存即无解除式，只有当拍判据）。
 * 码表     (Codes)      : 本件不占用任何全局数字码位。出口为 USINT 评分 + ENUM 分档 + BOOL，
 *                         数字码位待主控收口阶段统一派号（R46 码位规则）。
 * 红线自检 (Redline)    : R1 ✓ 零 GVL/VAR_EXTERNAL ｜ R2 ✓ 零 %I/%Q/%M ｜ R3 ✓ 纯 IEC 61131-3
 *                         R4 ✓ 除零前判零 + 浮点容差 ｜ R5 ✓ 声明逐行同行双语注释
 *                         R6 ✓ ENUM+CASE 含 ELSE ｜ R7 ✓ R_TRIG 段 0 无条件刷新
 * 修订历史 (Revision)   : 2026-11-19  v1.0.0  R46 首版（批次 1 · 序号 2）
 *==============================================================================*)

TYPE E_DL_EplGrade :
(
    eUnknown := 0,    // 本窗未评分（激励不足或组态非法） / Not scored this window
    eGood    := 10,   // 评分良好 / Score good
    eWatch   := 20,   // 评分关注（趋势劣化起点） / Score watch, degradation starting
    ePoor    := 30    // 评分劣化 / Score poor
);
END_TYPE

TYPE E_DL_EplState :
(
    eIdle := 0,    // 未取得首窗数据 / Awaiting first window
    eRun  := 10,   // 逐窗评分运行 / Scoring per window
    eBad  := 90    // 组态非法相（当拍可自愈） / Illegal configuration phase
);
END_TYPE

TYPE E_DL_EplCause :
(
    eNone       := 0,   // 无异常 / No anomaly
    eCfgIllegal := 1,   // 组态非法（分档线倒置/越界/比值下界非正） / Illegal configuration
    eNonFin     := 2,   // 期望值或下界非有限（NaN/Inf） / Non-finite expectation or floor
    eExcLow     := 3,   // 激励不足：期望脉冲数未过下界，本窗不评分 / Insufficient excitation, window not scored
    ePhaseBad   := 4    // 非法相位兜底 / Illegal phase fallback
);
END_TYPE

FUNCTION_BLOCK FB_DL_AxisEncoderPulseLostScore
VAR_INPUT
    nPulseCntWindow : DINT := 0;          // 窗内实测脉冲数（调用方累计，窗口起点清零） [cnt] / Measured pulses in window [cnt]
    fExpectWindow   : REAL := 0.0;        // 窗内期望脉冲数（|参考速度|×每毫米脉冲×窗长） [cnt] / Expected pulses in window [cnt]
    bWindowEnd      : BOOL := FALSE;      // 窗口结束触发，上升沿取一次快照 [-] / Window end trigger, snapshot on rising edge
    fRatioMin       : REAL := 0.01;       // 有效比值下界，域 > 0.0（防期望过小病态放大） [-] / Valid ratio lower bound, > 0.0
    nScoreGood      : INT := 98;          // 良好分档线，域 0..100 且 > nScoreWarn [分] / Good threshold, 0..100, > warn
    nScoreWarn      : INT := 90;          // 关注分档线，域 0..100 且 < nScoreGood [分] / Watch threshold, < good
    bReset          : BOOL := FALSE;      // 复位，上升沿回初始等待 [-] / Reset, rising edge returns to idle
END_VAR
VAR_OUTPUT
    fRatio  : REAL;                 // 本窗实测/期望比值（未评分时为 0.0） [-] / Measured over expected ratio this window
    nScore  : USINT;                // 本窗评分 0..100（未评分保持上窗值） [分] / Score 0..100, held when not scored
    eGrade  : E_DL_EplGrade;        // 评分分档出口 [-] / Score grade outlet
    bValid  : BOOL;                 // 本窗评分有效 [-] / Score valid this window
    bOverRun: BOOL;                 // 实测超期望（多脉冲，可能与丢脉冲相互掩盖） [-] / Pulses above expectation
    eState  : E_DL_EplState;        // 状态出口 [-] / State outlet
    eCause  : E_DL_EplCause;        // 本窗异常成因出口（信息级，当拍重算） [-] / Window anomaly cause, recomputed each scan
    bError  : BOOL;                 // 组态/输入非法标志（当拍重算，不锁存） [-] / Illegal config/input flag
END_VAR
VAR
    _eState  : E_DL_EplState := E_DL_EplState.eIdle;    // 内部相位（CASE 唯一写入目标） / Internal phase
    rtWin    : R_TRIG;              // 窗口结束沿实例，段 0 无条件调用 / Window-end edge instance
    rtReset  : R_TRIG;              // 复位沿实例，段 0 无条件调用 / Reset edge instance
    _nScore  : USINT;               // 评分锁存（未评分时保持） [分] / Held score
    _eCause  : E_DL_EplCause := E_DL_EplCause.eNone;   // 成因锁存前的当拍量（每拍重算） / Per-scan cause, recomputed
    _bNonFin : BOOL;                // 输入非有限当拍量 [-] / Non-finite input this scan
    _bCfgBad : BOOL;                // 组态非法当拍量 [-] / Illegal configuration this scan
    _bExcite : BOOL;                // 激励充足当拍量（期望值过下界） [-] / Sufficient excitation this scan
    _fRatio  : REAL;                // 当拍比值中间量 [-] / Ratio intermediate
END_VAR
VAR CONSTANT
    DL_EPL_EPS      : REAL := 1.0E-6;   // 浮点判零容差 [无量纲] / Float epsilon
    DL_EPL_SCORE_MAX: REAL := 100.0;    // 评分上限 [分] / Score ceiling
    DL_EPL_SCORE_MIN: REAL := 0.0;      // 评分下限 [分] / Score floor
END_VAR

(* —— 段 0：当拍量派生 + 沿实例无条件周期刷新 —— *)
_bNonFin := (fExpectWindow <> fExpectWindow) OR (fRatioMin <> fRatioMin);   // NaN 自反判 / NaN self-reflexive tests
_bCfgBad := (nScoreGood <= nScoreWarn) OR (nScoreGood > 100) OR (nScoreWarn < 0)   // 分档线几何闸 / Grade threshold geometry gate
         OR (nScoreWarn > 100) OR (fRatioMin <= 0.0) OR _bNonFin;                  // 比值下界闸 + 非有限 / Ratio floor and non-finite
_bExcite := (NOT _bNonFin) AND (fExpectWindow > DL_EPL_EPS)                 // 期望值须为正且有限 / Expectation must be positive and finite
         AND (fExpectWindow > (fRatioMin * DL_EPL_SCORE_MAX));              // 期望值下界 = 比值下界 × 100 脉冲口径 / Expectation floor in pulse counts
rtWin(CLK := bWindowEnd);                                                   // 窗口结束沿，每拍必调（R228A） / Window-end edge
rtReset(CLK := bReset);                                                     // 复位沿，每拍必调 / Reset edge

(* —— 段 1：单拍量预清零（锁存量 _nScore 不入清单，R107） —— *)
fRatio   := DL_EPL_SCORE_MIN;    // 比值每拍预清，评分分支同拍回填 / Ratio preset
nScore   := _nScore;             // 评分出口先回放锁存值，本窗有效时覆盖 / Score outlet replays held value
eGrade   := E_DL_EplGrade.eUnknown;   // 分档每拍预清 / Grade preset
eCause   := E_DL_EplCause.eNone;      // 成因每拍预清（信息级可重算，R189 例外条款） / Cause preset
bValid   := FALSE;               // 有效位每拍预清 / Validity preset
bOverRun := FALSE;               // 超发位每拍预清 / Over-run preset
bError   := FALSE;               // 非法标志每拍预清 / Error flag preset

(* —— 段 2：复位沿 —— *)
IF rtReset.Q THEN
    _eState := E_DL_EplState.eIdle;     // 回初始等首窗（无锁存故障，故只需相位复位） / Back to idle, no latch to clear
    _nScore := 0;                       // 评分锁存清零（复位是有意清历史） / Clear held score on explicit reset
END_IF

(* —— 段 3：组态/输入非法（当拍置位，不锁存；信息级不外溢为故障） —— *)
IF _bCfgBad THEN
    bError := TRUE;                     // 非法标志置位（同拍配对，R45） / Illegal flag set, same-scan pairing
    IF _bNonFin THEN
        eCause := E_DL_EplCause.eNonFin;    // 归因：输入非有限（优先于组态几何闸） / Cause: non-finite input, takes precedence
    ELSE
        eCause := E_DL_EplCause.eCfgIllegal;    // 归因：组态几何非法 / Cause: illegal configuration geometry
    END_IF
    _eState := E_DL_EplState.eBad;      // 入非法相（下拍自动回运行相） / Enter bad phase, self-heals next scan
END_IF

(* —— 段 4：窗口结束沿评分（单点写入评分锁存，避免同拍抹除，R187） —— *)
IF rtWin.Q AND (NOT _bCfgBad) THEN
    IF _bExcite THEN                                                          // 激励充足：真实评分 / Sufficient excitation: real scoring
        IF fExpectWindow > DL_EPL_EPS THEN                                    // 除零闸（双保险：_bExcite 已含下界） / Division guard
            _fRatio := INT_TO_REAL(nPulseCntWindow) / fExpectWindow;          // 实测 / 期望 / Measured over expected
        ELSE
            _fRatio := DL_EPL_SCORE_MIN;                                      // 病态期望值：比值记 0 / Degenerate expectation: ratio zero
        END_IF
        fRatio := _fRatio;                                                    // 比值出口（本窗有效值） / Ratio outlet for a valid window
        IF _fRatio >= 1.0 THEN                                                // 达到或超过期望 / At or above expectation
            _nScore := 100;                                                   // 满分封顶（超发不奖分） / Ceiling at full score
            bOverRun := _fRatio > 1.02;                                       // 超发 2% 以上给提示（防双向掩盖） / Over-run hint above 2 percent
        ELSE
            IF _fRatio < DL_EPL_SCORE_MIN THEN
                _fRatio := DL_EPL_SCORE_MIN;                                  // 负计数（脏数据）钳到下限 / Clamp dirty negative count
            END_IF
            _nScore := REAL_TO_USINT(_fRatio * DL_EPL_SCORE_MAX);             // 线性折分 0..100 / Linear score scaling
        END_IF
        IF _nScore > 100 THEN
            _nScore := 100;                                                   // 类型上限再兜一层（USINT 溢出前置） / Second ceiling before USINT range
        END_IF
        bValid := TRUE;                                                       // 本窗评分有效 / Window scored
        nScore := _nScore;                                                    // 评分出口与锁存同源 / Score outlet from latch
    ELSE
        bValid := FALSE;                                                      // 激励不足：本窗不评分（禁记 100 分） / No excitation: no scoring, never 100
        eCause := E_DL_EplCause.eExcLow;                                      // 归因：激励不足（与本窗不评分同因） / Cause: insufficient excitation
    END_IF
END_IF

(* —— 段 5：分档映射（与 nScale 同源，出口单点） —— *)
IF bValid THEN
    IF INT_TO_USINT(nScoreGood) <= nScore THEN
        eGrade := E_DL_EplGrade.eGood;         // 良好档 / Good grade
    ELSIF INT_TO_USINT(nScoreWarn) <= nScore THEN
        eGrade := E_DL_EplGrade.eWatch;        // 关注档 / Watch grade
    ELSE
        eGrade := E_DL_EplGrade.ePoor;         // 劣化档 / Poor grade
    END_IF
ELSE
    eGrade := E_DL_EplGrade.eUnknown;          // 未评分档 / Unknown grade
END_IF

(* —— 段 6：相位机（ENUM 全成员显式标签 + ELSE 兜底，R128） —— *)
CASE _eState OF

E_DL_EplState.eIdle:
    IF (NOT _bCfgBad) AND (rtWin.Q OR _bExcite) THEN    // 出口 1：组态合法且已来窗/已见激励 / Legal config and a window seen
        _eState := E_DL_EplState.eRun;
    ELSIF _bCfgBad THEN                                 // 出口 2：组态非法 / Illegal configuration
        _eState := E_DL_EplState.eBad;
    END_IF

E_DL_EplState.eRun:
    IF _bCfgBad THEN                                    // 出口 1：组态转非法 / Configuration went illegal
        _eState := E_DL_EplState.eBad;
    ELSIF rtReset.Q THEN                                // 出口 2：复位回等首窗 / Reset back to first window
        _eState := E_DL_EplState.eIdle;
    END_IF

E_DL_EplState.eBad:
    IF NOT _bCfgBad THEN                                // 出口：组态恢复即自愈回运行 / Self-heal once configuration is legal
        _eState := E_DL_EplState.eRun;
    END_IF

ELSE
    bError  := TRUE;                                    // 非法相位兜底：置非法标志 / Illegal-phase fallback flag
    eCause  := E_DL_EplCause.ePhaseBad;                 // 归因：非法相位 / Cause: illegal phase
    _eState := E_DL_EplState.eBad;                      // 强拉非法相 / Force bad phase

END_CASE

eState := _eState;                                      // 状态出口 / State outlet

END_FUNCTION_BLOCK

(* ---- FB_DL_AxisFollowErrGuard.st ---- *)
(*
  FB_DL_AxisFollowErrGuard  —  轴跟随误差窗口监视 / Axis following-error window guard
  分类 Category : DL_Motion
  版本 Version  : 1.0.0
  来源 Source   : t1-6-plcopen — 运动守卫族零检索深化（P0-1 解除式教训落地）
  溯源 Origin   : clean-room 实现，PLCopen 跟随误差监视语义公开借鉴，未复制任何源码行
  功能 Function : 1) 经 I_DL_MotionAxis 读 fPosition（当拍量），与注入的位置指令 fPosSet
                  做差得跟随误差；|fVelocity| > fVelGate（运动门控）且误差 > fErrBand
                  持续 tErrTo → 故障级 03A9 锁存；
                  2) 误差进入 80% 带置预警沿信息级 04A8；误差回带内置恢复信息级 04A9；
                  3) 故障解除式全当拍量（R240 落地）：rtReset.Q AND NOT iAxis.bError
                  AND 误差回带内，逐 BOOL 标注见段 4；
                  4) 非有限误差 → 故障级 03AA 防御兜底锁存。
  边界 Boundary : ① I_DL_MotionAxis 无 fPosSet 属性（接口实测），位置指令由调用方引脚注入，
                  本件不实例化轴实现块；
                  ② 组态闸：fErrBand <= 0 或超时 <= 0 或门速 < 0 → 03A8 锁存；
                  ③ 门速 fVelGate = 0 语义为「静止也判」，显式允许（下移 0.0 语义合法）；
                  ④ 无 GVL 依赖：纯引脚输入输出，无外部变量引用，无物理 IO 地址。
  依赖 Depends  : I_DL_MotionAxis（注入，不实例化）；Standard.library（TON / R_TRIG）
  码表 Error codes（Motion 段 0004，窗口 03A8~03AA / 04A8~04AA）:
    16#0004_03A8 故障级：组态非法（误差带/超时/门速域非法），锁存至 bReset
    16#0004_03A9 故障级：跟随误差超窗（运动门控下持续 tErrTo），锁存至 bReset
    16#0004_03AA 故障级：跟随误差非有限（防御兜底），锁存至 bReset
    16#0004_04A8 信息级：超窗预警沿（误差进入 80% 带）
    16#0004_04A9 信息级：误差恢复正常沿（回带内）
    16#0004_04AA 信息级：守卫使能沿（bEnable 上升沿）
  修订历史 Revision :
    2026-11-19  v1.0.0  R41 首版（批次 2 · 序号 4）
*)

FUNCTION_BLOCK FB_DL_AxisFollowErrGuard
VAR_INPUT
    fPosSet      : REAL := 0.0;       // 位置指令 [mm 或 deg]，调用方注入 / Position command injected by caller
    fErrBand     : REAL := 0.5;       // 跟随误差带半宽 [mm 或 deg]，域 >= 0 / Following-error band half width
    fVelGate     : REAL := 1.0;       // 运动门速 [mm/s]，域 >= 0，0 = 静止也判 / Motion gating speed
    tErrTo       : TIME := T#500MS;   // 超窗确认超时 [ms]，域 > 0 / Over-window confirm timeout
    bEnable      : BOOL := FALSE;     // 守卫使能 [-] / Guard enable
    bReset       : BOOL := FALSE;     // 复位，上升沿清故障锁存 / Reset edge clears fault latch
END_VAR
VAR_IN_OUT
    iAxis        : I_DL_MotionAxis;   // 运动轴引用（注入，不实例化）/ Motion axis reference
END_VAR
VAR_OUTPUT
    fFollowErr   : REAL;              // 跟随误差绝对值 [mm 或 deg] / Absolute following error
    bWarn        : BOOL;              // 预警标志（误差 > 80% 带）/ Warning flag
    bFault       : BOOL;              // 故障锁存标志 / Fault latch flag
    bError       : BOOL;              // 故障级标志（与锁存位同源）/ Fault flag
    nErrId       : UDINT;             // 事件码，0 = 无事件 / Event code
END_VAR
VAR
    tonErrTo     : TON;               // 超窗确认定时器，无条件周期刷新 / Over-window confirm timer
    rtReset      : R_TRIG;            // 复位沿实例，无条件刷新 / Reset edge instance
    rtEn         : R_TRIG;            // 使能沿实例，无条件刷新 / Enable edge instance
    _fErr        : REAL;              // 跟随误差中间量 [mm 或 deg] / Following error intermediate
    _bFault      : BOOL;              // 故障锁存位（锁存量）/ Latched fault bit
    _uFault      : UDINT;             // 故障码锁存（锁存量）/ Latched fault code
    _uInfo       : UDINT;             // 信息码，每拍重算 / Transient info code
    _bWarnPrev   : BOOL;              // 上拍预警镜像（预警沿判据）/ Previous warn mirror
    _bInBandPrev : BOOL;              // 上拍带内镜像（恢复沿判据）/ Previous in-band mirror
END_VAR

(* —— 段 0：定时器与沿实例无条件周期刷新（禁置于 IF/CASE 内） —— *)
_fErr := ABS(fPosSet - iAxis.fPosition);              // 跟随误差（全当拍量）
rtReset(CLK := bReset);                               // 复位沿（每拍必调）
rtEn(CLK := bEnable);                                 // 使能沿（每拍必调）
tonErrTo(IN := bEnable AND (ABS(iAxis.fVelocity) > fVelGate) AND (_fErr > fErrBand), PT := tErrTo);
                                                      // 超窗确认（运动门控，每拍必调）

(* —— 段 1：单拍量预清零（锁存量 _bFault/_uFault 不入清单，禁同拍抹除） —— *)
_uInfo := 16#0000_0000;             // 信息码每拍重算
bWarn := FALSE;                     // 预警出口缺省 FALSE
nErrId := 16#0000_0000;             // 事件码缺省无事件

(* —— 段 2：复位沿 + 组态域闸（当拍量判据） —— *)
IF rtReset.Q THEN                   // rtReset.Q = 当拍量
    _bFault := FALSE;               // 清故障锁存位
    _uFault := 16#0000_0000;        // 清故障锁存码
END_IF
IF (fErrBand < 0.0) OR (fVelGate < 0.0) OR (TIME_TO_DINT(tErrTo) <= 0) THEN
    _uFault := 16#0004_03A8;        // 故障级：组态非法
    _bFault := TRUE;
END_IF

(* —— 段 3：非有限误差防御兜底（NaN 自反判，禁近似阈值） —— *)
IF (_fErr <> _fErr) OR ((_fErr - _fErr) <> (_fErr - _fErr)) THEN
    _uFault := 16#0004_03AA;        // 故障级：误差非有限
    _bFault := TRUE;
    _fErr := 0.0;                   // 出口安全侧归零
END_IF

(* —— 段 4：故障聚合与超窗锁存（判据全当拍量） —— *)
IF (NOT _bFault) AND tonErrTo.Q THEN
    _uFault := 16#0004_03A9;        // 故障级：跟随误差超窗锁存
    _bFault := TRUE;
END_IF

(* —— 段 5：故障解除式（R240 落地，逐 BOOL 标注）：
     rtReset.Q = 当拍量；iAxis.bError = 当拍量；(_fErr <= fErrBand) = 当拍量。
     三者均不含锁存量（_bFault/_uFault），解除边真实可达。 —— *)
IF rtReset.Q AND (NOT iAxis.bError) AND (_fErr <= fErrBand) THEN
    _bFault := FALSE;               // 清故障锁存位（锁存量，仅此当拍量解除沿可清）
    _uFault := 16#0000_0000;        // 清故障锁存码（锁存量，同上唯一解除路径）
END_IF

(* —— 段 6：预警与信息码派生（当拍量判据） —— *)
IF (NOT _bFault) AND bEnable THEN
    bWarn := _fErr > (fErrBand * 0.8);      // 预警：误差进入 80% 带
    IF bWarn AND (NOT _bWarnPrev) THEN
        _uInfo := 16#0004_04A8;             // 信息级：预警沿
    END_IF
    IF (NOT bWarn) AND _bInBandPrev AND (NOT _bWarnPrev) THEN
        _uInfo := 16#0004_04A9;             // 信息级：误差恢复沿（带内持续）
    END_IF
END_IF
IF rtEn.Q THEN
    _uInfo := 16#0004_04AA;         // 信息级：使能沿（覆盖预警沿，使能优先报告）
END_IF

(* —— 段 7：出口单点映射（锁存码回放，禁同拍抹除） —— *)
fFollowErr := _fErr;                // 误差出口镜像
IF _bFault THEN
    nErrId := _uFault;              // 故障锁存码回放
    bWarn := FALSE;                 // 故障期预警强制 FALSE（安全侧）
ELSE
    nErrId := _uInfo;               // 信息码
END_IF
bFault := _bFault;                  // 锁存位出口
bError := _bFault;                  // 故障标志与锁存位同源
_bWarnPrev := bWarn;                // 预警沿判据快照
_bInBandPrev := (NOT bWarn);        // 带内镜像快照

END_FUNCTION_BLOCK

(* ---- FB_DL_AxisFollowingErrorMonitor.st ---- *)
(*
    FB_DL_AxisFollowingErrorMonitor —— 跟随误差监视
    ------------------------------------------------------------------
    分类      : DL_Motion / Monitor
    前缀      : FB_DL_
    版本      : 1.0.0
    溯源      : T1-6 PLCopen（只借「跟随误差监视属运动控制监视功能」的公开语义，
                不自造轴状态机）；T2-4 监视参数域为次源；
                确认窗、静止带、阈值交换逻辑与码位 100% 自有；clean-room 重写，
                未复制任何闭源厂商源码，参考实现仅限 MIT/Apache 许可
    平台      : 纯 IEC 61131-3，CODESYS V3.5+ / TwinCAT 3 / InoProShop 通用
    作者      : 道莅代码库 · PLC编程专家（R18）
    ------------------------------------------------------------------
    功能说明  : 消费「指令位置 + 实际位置」两个快照，算跟随误差并做三级判定
                （正常 / 预警 / 故障），带确认时间与静止带豁免；
                本件不自造轴状态、不发运动指令——轴状态唯一属主在 FB_DL_SingleAxis，
                本件只是被动消费者（同 PassiveHomingMonitor 纪律）；
                阈值倒置自动交换而不是报故障：现场参数填反极常见，直接锁死会停线；
                静止带内误差视为正常并清计时，防静止噪声误跳；
                eErr（参数 / 信号类）与 bFault（工艺跟随超差）分开出口，便于 HMI 分组。
    错误码    : 16#0004_01C7 阈值倒置已自动交换 / 阈值超域已钳位——信息级，不置故障
                16#0004_01C8 预留禁用（信息级，不得挪用）
                16#0004_02D5 位置快照非有限（NaN / 正负 INF）——故障级，判定冻结
                16#0004_02D6 越限持续超确认窗（与 bFault 同拍置位，可追溯标识）——故障级
                16#0004_02D7 预留禁用（故障级，不得挪用）
    码位总账  : 16#0004_01C7 用 / 16#0004_01C8 预留 ｜ 16#0004_02D5 用 / 16#0004_02D6 用 / 16#0004_02D7 预留
    状态机    : 无 CASE，判定由两个 TON 与一个故障锁存位承载，非法状态不可能出现
    采样约定  : fbTrigReset 与两个 TON 在本体首部无条件调用；静止时只把定时器 IN 引脚
                置 FALSE，绝不把 TON 调用放进 IF（否则 ET 冻结产生幽灵确认）。
    修订记录  : 2026-11-16 v1.0.0 首次入库（R18）
*)
FUNCTION_BLOCK FB_DL_AxisFollowingErrorMonitor
VAR_INPUT
    bEnable         : BOOL;                    // 使能，FALSE 清判定并按正常输出 / enable, FALSE clears the verdict and reports normal
    bReset          : BOOL;                    // 复位，上升沿清故障与计时 / reset, rising edge clears the fault and the timers
    fSetPosition    : REAL := 0.0;             // 指令位置，由运动层注入 [mm] / commanded position injected by the motion layer [mm]
    fActPosition    : REAL := 0.0;             // 实际位置反馈 [mm] / actual position feedback [mm]
    fWarnLimit      : REAL := 0.5;             // 预警阈值，必须大于 0 [mm] / warning threshold, must exceed zero [mm]
    fFaultLimit     : REAL := 2.0;             // 故障阈值，必须大于 0 且大于预警阈值 [mm] / fault threshold, must exceed zero and the warning threshold [mm]
    tConfirmTime    : TIME := T#200MS;         // 越限持续确认时间，0 = 立即判定 [ms] / over-limit confirmation time, 0 = immediate [ms]
    fStandstillBand : REAL := 0.05;            // 静止带，误差在此内视为正常（噪声容忍）[mm] / standstill band, the error inside it counts as normal [mm]
    bInMotion       : BOOL := FALSE;           // 运动中标志，FALSE 时确认时间不累加 / in-motion flag, the timers do not accumulate when FALSE
END_VAR
VAR_OUTPUT
    fError    : REAL;                          // 跟随误差（指令减实际）[mm] / following error, command minus actual [mm]
    fErrorAbs : REAL;                          // 误差绝对值 [mm] / absolute following error [mm]
    bWarn     : BOOL;                          // 预警（越预警阈值超确认时间）/ warning, over the warning threshold beyond the confirmation time
    bFault    : BOOL;                          // 故障（越故障阈值超确认时间，已锁存）/ fault, over the fault threshold beyond the confirmation time, latched
    tOverTime : TIME;                          // 当前越预警阈值已持续时间 [ms] / time spent above the warning threshold [ms]
    eErr      : UDINT;                         // 错误码（参数 / 信号类），0=正常 / error id of the parameter or signal class, 0=ok
    bError    : BOOL;                          // 故障标志（参数类），与 bFault 区分 / error flag of the parameter class, distinct from bFault
END_VAR
VAR
    fbTrigReset   : R_TRIG;                    // 复位沿检测实例，本体首部无条件刷新 / reset edge instance, refreshed unconditionally
    fbConfirmWarn : TON;                       // 预警确认定时器，本体首部无条件刷新 / warning confirmation timer, refreshed unconditionally
    fbConfirmFault: TON;                       // 故障确认定时器，本体首部无条件刷新 / fault confirmation timer, refreshed unconditionally
    fWarnEff      : REAL;                      // 生效预警阈值，交换与钳位后 [mm] / effective warning threshold after swap and clamp [mm]
    fFaultEff     : REAL;                      // 生效故障阈值，交换与钳位后 [mm] / effective fault threshold after swap and clamp [mm]
    fTmpSwap      : REAL;                      // 阈值交换中间量 [mm] / threshold swap intermediate [mm]
    fErrorLast    : REAL;                      // 末次有效误差，非有限时保持 [mm] / last valid error held through non-finite cycles [mm]
    bFaultLatch   : BOOL;                      // 故障锁存位，仅复位清除 / fault latch, cleared by reset only
    bFrozen       : BOOL;                      // 判定冻结标志，快照非有限时为 TRUE / verdict freeze flag, TRUE on a non-finite snapshot
    bNonFin       : BOOL;                      // 快照非有限判定标志 / snapshot non-finite flag
END_VAR
VAR CONSTANT
    DL_FE_MIN_LIMIT  : REAL := 0.001;          // 阈值下限 [mm] / threshold lower bound [mm]
    DL_FE_MAX_LIMIT  : REAL := 1.0E4;          // 阈值上限 [mm] / threshold upper bound [mm]
    DL_FE_INF_GUARD  : REAL := 4.0E38;         // 非有限幅值判定阈值 [mm] / non-finite magnitude guard [mm]
    DL_FLOAT_EPS     : REAL := 1.0E-6;         // 浮点判等容差 [mm] / float equality tolerance [mm]
    DL_FE_ZERO       : REAL := 0.0;            // 零值常量，避免裸字面量 [无量纲] / zero constant, avoids a bare literal [dimensionless]
    DL_FE_ONE        : REAL := 1.0;            // 一值常量，用于交换判据 [无量纲] / one constant used by the swap criterion [dimensionless]
END_VAR

// 段 1｜边沿实例无条件周期刷新（红线：严禁放入条件分支）/ segment 1, unconditional edge refresh
fbTrigReset(CLK := bReset);

// 段 2｜输出与错误状态预置 / segment 2, preset outputs and error status
eErr := 0;                                     // 预置无错误 / preset no error
bError := FALSE;                               // 预置无故障标志 / preset no error flag
bWarn := FALSE;                                // 预置无预警 / preset no warning
bFrozen := FALSE;                              // 预置不冻结 / preset not frozen

// 段 3｜失能期的记忆与锁存清理：本件无首扫专用初值，状态由 bFaultLatch 与 fErrorLast 承载 / segment 3, memory and latch clearing while disabled, no dedicated first-scan init needed
IF NOT bEnable THEN
    fErrorLast := DL_FE_ZERO;                  // 失能清误差记忆 / clear the error memory while disabled
    bFaultLatch := FALSE;                      // 失能清故障锁存 / clear the fault latch while disabled
END_IF

// 段 4｜阈值域校正：先钳位再判倒置，倒置自动交换（信息级，绝不锁死生产）/ segment 4, threshold correction
fWarnEff := MIN(MAX(fWarnLimit, DL_FE_MIN_LIMIT), DL_FE_MAX_LIMIT);   // 预警阈值双侧钳位 / clamp the warning threshold both sides
fFaultEff := MIN(MAX(fFaultLimit, DL_FE_MIN_LIMIT), DL_FE_MAX_LIMIT); // 故障阈值双侧钳位 / clamp the fault threshold both sides
IF ABS(fWarnEff - fWarnLimit) > DL_FLOAT_EPS THEN
    eErr := 16#0004_01C7;                      // 钳位提示（信息级不置故障）/ clamp hint, info level never raises a fault
END_IF
IF ABS(fFaultEff - fFaultLimit) > DL_FLOAT_EPS THEN
    eErr := 16#0004_01C7;                      // 钳位提示（信息级不置故障）/ clamp hint, info level never raises a fault
END_IF
IF fWarnEff >= fFaultEff THEN
    fTmpSwap := fWarnEff;                      // 暂存预警阈值 / hold the warning threshold
    fWarnEff := fFaultEff;                     // 交换下限 / swap the lower bound
    fFaultEff := fTmpSwap;                     // 交换上限 / swap the upper bound
    eErr := 16#0004_01C7;                      // 交换提示（信息级不置故障）/ swap hint, info level never raises a fault
END_IF

// 段 5｜误差计算与非有限闸：非有限时保持末次有效误差并冻结判定 / segment 5, error computation and non-finite gate
bNonFin := (fSetPosition <> fSetPosition)
        OR (fSetPosition > DL_FE_INF_GUARD) OR (fSetPosition < -DL_FE_INF_GUARD)
        OR (fActPosition <> fActPosition)
        OR (fActPosition > DL_FE_INF_GUARD) OR (fActPosition < -DL_FE_INF_GUARD); // 双快照同口径检查 / both snapshots checked the same way
IF bNonFin THEN
    eErr := 16#0004_02D5;                      // 快照非有限故障码 / non-finite snapshot fault id
    bError := TRUE;                            // 置故障标志 / raise the error flag
    fError := fErrorLast;                      // 保持末次有效误差 / hold the last valid error
    bFrozen := TRUE;                           // 冻结判定与计时 / freeze the verdict and the timers
ELSE
    fError := fSetPosition - fActPosition;     // 指令减实际 / command minus actual
    fErrorLast := fError;                      // 刷新误差记忆 / refresh the error memory
END_IF
fErrorAbs := ABS(fError);                      // 绝对值出口 / absolute value output

// 段 6｜静止带豁免：带内视为正常且清计时（不改定时器调用位置，只改 IN 引脚）/ segment 6, standstill band exemption
IF fErrorAbs <= fStandstillBand THEN
    bFrozen := TRUE;                           // 静止带内冻结计时，防噪声误跳 / freeze the timers inside the band, prevents noise trips
END_IF

// 段 7｜定时器每拍调用一次且位于条件分支之外，IN 引脚承载全部条件 / segment 7, one call per cycle outside any branch, the IN pin carries every condition
fbConfirmWarn(IN := bEnable AND (NOT bFrozen) AND bInMotion AND (fErrorAbs > fWarnEff), PT := tConfirmTime);
fbConfirmFault(IN := bEnable AND (NOT bFrozen) AND bInMotion AND (fErrorAbs > fFaultEff), PT := tConfirmTime);

// 段 8｜复位沿清故障与计时（优先于判定）/ segment 8, reset clears the fault and the timers
IF fbTrigReset.Q THEN
    bFaultLatch := FALSE;                      // 清故障锁存 / clear the fault latch
    bWarn := FALSE;                            // 清预警 / clear the warning
END_IF

// 段 9｜判定：故障优先于预警，故障锁存后只能复位清除 / segment 9, verdict with the fault taking priority
IF fbConfirmFault.Q THEN
    bFaultLatch := TRUE;                       // 越故障阈值超确认窗，锁存 / above the fault threshold beyond the confirmation time, latch it
    eErr := 16#0004_02D6;                      // 越限持续故障码，与 bFault 同拍置位 / over-limit sustained fault id, set on the same cycle as bFault
    bError := TRUE;                            // 置故障标志，便于 HMI 与 bFault 同屏追溯 / raise the error flag so the HMI can trail both flags together
END_IF
IF (NOT bFaultLatch) AND fbConfirmWarn.Q THEN
    bWarn := TRUE;                             // 越预警阈值超确认窗 / above the warning threshold beyond the confirmation time
END_IF

// 段 10｜输出 / segment 10, publish the outputs
bFault := bFaultLatch;                         // 工艺故障出口 / process fault output
tOverTime := fbConfirmWarn.ET;                 // 越限已持续时间取预警定时器 ET / the elapsed time comes from the warning timer
IF bFaultLatch THEN
    bWarn := FALSE;                            // 故障优先，预警让位 / the fault takes priority, the warning steps aside
END_IF
IF NOT bEnable THEN
    bFault := FALSE;                           // 失能即按正常输出 / disabled reports normal
    bWarn := FALSE;                            // 失能即无预警 / no warning while disabled
    tOverTime := T#0MS;                        // 计时清零 / clear the elapsed time
END_IF
END_FUNCTION_BLOCK

(* ---- FB_DL_AxisFrictionFf.st ---- *)
(*
  组件名 Component   : FB_DL_AxisFrictionFf
  子库 Sublibrary    : DL_Motion
  版本 Version       : 1.0.0
  兼容性 Platform    : CODESYS 3.5 / TwinCAT 3 / 汇川 InoProShop / Machine Expert（仅 Standard.library）
  功能 Function      : 摩擦转矩前馈：
                       1) 静/动摩擦分段：|速度| < 静动切换阈 → 静摩擦段（出全静摩擦值），
                       否则动摩擦段（出动摩擦值）；
                       2) 速度方向切换滞环：方向电平只在速度越过零速迟滞带后翻转，
                       防零速附近前馈符号抖动；
                       3) 前馈系数钳位：fFfGain 域 [0, 1]，域外钳位并告警锁存；
                       4) 分段切换与换向均经一阶惯性平滑（tSmooth），防前馈阶跃。
  边界 Boundary      : ① 本件只出前馈转矩，不参与闭环（叠加由上层转矩合成）；
                       ② 组态闸：静摩擦 < 动摩擦（物理不可能）、系数负值、tCycle 零 → 故障；
                       ③ 非有限值（NaN 自反 + 无穷差值自减）判输入非法锁存；
                       ④ 故障锁存解除唯一路径 = bReset 上升沿（输入引脚，恒可达）；
                       ⑤ 无全局变量引用、无外部变量声明、无物理地址寻址。
  依赖 Depends       : Standard.library（R_TRIG）
  溯源 Origin        : 道莅自研 clean-room（参考 t2-4-s7-motion 前馈分类与参数域，
                       零代码行复制）
  码位 Code          : 16#04_0_AB
  码表 Error codes（Motion 格 04_0_AB，单轨：故障 0x02AB / 信息 0x01AB）:
    16#0004_02AB 故障级：组态非法（静摩擦 < 动摩擦 / 系数负 / tCycle 零）或输入
                 非有限，锁存至 bReset 上升沿
    16#0004_01AB 信息级：前馈系数已钳位（域 [0,1] 越界当拍，瞬时口径）
  修订历史 Revision  :
    2026-11-19  v1.0.0  R44 首版（批次 2 · 序号 8）
*)

TYPE E_DL_AffState :
(
    eIdle  := 0,    // 空闲：未使能，前馈归零 / Idle, feedforward zeroed
    eRun   := 10,   // 运行：分段前馈 / Running, segmented feedforward
    eFault := 90    // 故障：组态/输入锁存 / Fault, latched
);
END_TYPE

TYPE E_DL_AffZone :
(
    eStatic := 0,   // 静摩擦段：|速度| < 切换阈 / Static zone
    eDynamic := 10, // 动摩擦段：|速度| >= 切换阈 / Dynamic zone
    eHold   := 20   // 保持段：故障相冻结 / Hold zone, fault frozen
);
END_TYPE

FUNCTION_BLOCK FB_DL_AxisFrictionFf
VAR_INPUT
    bEnable      : BOOL;                   // 使能（电平）[-] / Enable
    bReset       : BOOL;                   // 上升沿清故障锁存 [-] / Reset edge
    fVelCmdMmS   : REAL;                   // 速度指令 [mm/s]，符号即方向 / Velocity command
    fFricStaticNm: REAL := 2.0;            // 静摩擦幅值 [牛·米] / Static friction magnitude
    fFricDynNm   : REAL := 1.0;            // 动摩擦幅值 [牛·米] / Dynamic friction magnitude
    fSwitchVelMmS: REAL := 2.0;            // 静动切换速度阈 [mm/s] / Static-dynamic switch threshold
    fHystVelMmS  : REAL := 0.5;            // 换向迟滞带 [mm/s] / Direction hysteresis band
    fFfGain      : REAL := 1.0;            // 前馈系数 [无量纲]，域 0..1 / Feedforward gain
    tSmooth      : TIME := T#100MS;        // 分段/换向平滑惯性 [毫秒] / Smoothing lag
    tCycle       : TIME := T#10MS;         // 扫描周期 [毫秒] / Scan cycle time
END_VAR
VAR_OUTPUT
    fFfTorqueNm  : REAL;                   // 前馈转矩输出 [牛·米] / Feedforward torque
    eFricZone    : E_DL_AffZone;           // 当前摩擦段出口 / Friction zone outlet
    bGainClamped : BOOL;                   // 系数已钳位标志 [-] / Gain clamped flag
    eState       : E_DL_AffState;          // 状态出口，段尾单点映射 / State outlet
    bError       : BOOL;                   // 故障锁存标志 [-] / Fault latch flag
    uErrId       : UDINT;                  // 事件码，0 = 无事件 / Event code
END_VAR
VAR
    rtReset : R_TRIG;                      // 复位沿实例，段 0 无条件刷新 / Reset edge
    _eState : E_DL_AffState := E_DL_AffState.eIdle;    // 内部相位（CASE 唯一写入目标）/ Internal phase
    _bDirPos: BOOL;                        // 方向电平（迟滞后）[-] / Direction level
    _bDirSeen: BOOL;                       // 首方向已建立标志 [-] / First direction established
    _fDemand: REAL;                        // 平滑前前馈需求 [牛·米] / Pre-smooth demand
    _fSmK   : REAL;                        // 平滑系数 [无量纲] / Smoothing coefficient
    _fGainUse: REAL;                       // 生效前馈系数 [无量纲] / Effective gain
    _eZone  : E_DL_AffZone := E_DL_AffZone.eStatic;    // 内部段（CASE 唯一写入目标）/ Internal zone
    _bFault : BOOL;                        // 故障锁存位（锁存量） / Latched fault bit
    _uFault : UDINT;                       // 故障码锁存（锁存量） / Latched fault code
    _bCfgBad: BOOL;                        // 组态非法当拍量 [-] / Config illegal flag
    _bNonFin: BOOL;                        // 输入非有限当拍量 [-] / Non-finite input flag
END_VAR
VAR CONSTANT
    DL_GAIN_MAX : REAL := 1.0;             // 前馈系数上限 [无量纲] / Gain ceiling
    DL_ZERO     : REAL := 0.0;             // 零常量 [工程单位] / Zero constant
    DL_ONE      : REAL := 1.0;             // 单位常量 [无量纲] / Unity constant
    DL_ABS_MAX  : REAL := 1.0E30;          // 有限值判定上界 [工程单位] / Finite bound
    DL_MS_PER_S : REAL := 1000.0;          // 毫秒 → 秒换算系数 [毫秒/秒] / Milliseconds per second
END_VAR

(* —— 段 0｜沿实例每拍无条件刷新（禁置于 IF/CASE 内） —— *)
rtReset(CLK := bReset);

(* —— 段 1｜瞬时量预清零（锁存量 _bFault/_uFault/_bDirSeen/_fFfTorqueNm 不入清单） —— *)
uErrId   := 16#0000_0000;
bGainClamped := FALSE;
_bCfgBad := FALSE;
_bNonFin := FALSE;

(* —— 段 2｜复位沿：故障一次性清干净，相位回空闲，前馈归零 —— *)
IF rtReset.Q THEN
    _bFault := FALSE;
    _uFault := 16#0000_0000;
    fFfTorqueNm := DL_ZERO;
    _eState := E_DL_AffState.eIdle;
END_IF

(* —— 段 3｜组态闸与非有限判据（覆盖全部参与换算引脚） —— *)
IF (fFricStaticNm < fFricDynNm) OR (fFricStaticNm < DL_ZERO) OR (fFricDynNm < DL_ZERO)
   OR (fFfGain < DL_ZERO) OR (fSwitchVelMmS <= DL_ZERO) OR (fHystVelMmS <= DL_ZERO)
   OR (tCycle = T#0S) THEN
    _bCfgBad := TRUE;
END_IF
IF (fVelCmdMmS <> fVelCmdMmS) OR ((fVelCmdMmS - fVelCmdMmS) <> DL_ZERO) THEN
    _bNonFin := TRUE;
END_IF

(* —— 段 4｜主状态机：三态全覆盖 + ELSE 兜底 —— *)
CASE _eState OF

E_DL_AffState.eIdle:
    IF bEnable AND (NOT _bCfgBad) AND (NOT _bNonFin) THEN
        _bDirSeen := FALSE;
        _bDirPos  := FALSE;
        fFfTorqueNm := DL_ZERO;
        _eState := E_DL_AffState.eRun;
    ELSIF bEnable AND (_bCfgBad OR _bNonFin) THEN
        _bFault := TRUE;
        _uFault := 16#0004_02AB;
        bError  := TRUE;
        _eState := E_DL_AffState.eFault;
    END_IF

E_DL_AffState.eRun:
    IF NOT bEnable THEN
        fFfTorqueNm := DL_ZERO;
        _eState := E_DL_AffState.eIdle;  // 使能撤销回空闲，前馈归零
    ELSIF _bNonFin THEN
        _bFault := TRUE;                 // 运行中输入非有限：锁存
        _uFault := 16#0004_02AB;
        bError  := TRUE;
        _eState := E_DL_AffState.eFault;
    ELSE
        (* 前馈系数钳位：域 [0,1]，越界钳位并留信息码 *)
        _fGainUse := fFfGain;
        IF _fGainUse > DL_GAIN_MAX THEN
            _fGainUse := DL_GAIN_MAX;
            bGainClamped := TRUE;
            uErrId := 16#0004_01AB;      // 信息级：系数钳位（瞬时口径）
        END_IF
        (* 方向迟滞：越零速迟滞带才翻转，防符号抖动 *)
        IF (NOT _bDirPos) AND (fVelCmdMmS > fHystVelMmS) THEN
            _bDirPos := TRUE;
            _bDirSeen := TRUE;
        ELSIF _bDirPos AND (fVelCmdMmS < -fHystVelMmS) THEN
            _bDirPos := FALSE;
            _bDirSeen := TRUE;
        END_IF
        (* 静/动分段 + 符号合成 *)
        IF ABS(fVelCmdMmS) < fSwitchVelMmS THEN
            _eZone := E_DL_AffZone.eStatic;
            IF _bDirPos THEN
                _fDemand := fFricStaticNm;
            ELSE
                _fDemand := -fFricStaticNm;
            END_IF
        ELSE
            _eZone := E_DL_AffZone.eDynamic;
            IF _bDirPos THEN
                _fDemand := fFricDynNm;
            ELSE
                _fDemand := -fFricDynNm;
            END_IF
        END_IF
        IF NOT _bDirSeen THEN
            _fDemand := DL_ZERO;         // 首方向未建立：需求归零
        END_IF
        _fDemand := _fDemand * _fGainUse;
        (* 一阶惯性平滑：tSmooth 零时直通 *)
        IF tSmooth = T#0S THEN
            _fSmK := DL_ONE;
        ELSE
            _fSmK := (TIME_TO_REAL(tCycle) / DL_MS_PER_S)
                     / ((TIME_TO_REAL(tCycle) / DL_MS_PER_S)
                        + TIME_TO_REAL(tSmooth) / DL_MS_PER_S);
        END_IF
        fFfTorqueNm := fFfTorqueNm + _fSmK * (_fDemand - fFfTorqueNm);
    END_IF

E_DL_AffState.eFault:
    bError := TRUE;                      // 故障相驻留：前馈冻结保持，只认复位沿（段 2 迁出）
    ;                                    // （冻结语义：fFfTorqueNm 保持最后值，禁降级归零不声明）
    _eZone := E_DL_AffZone.eHold;        // 段出口进保持段（名实双出口）

ELSE
    _bFault := TRUE;                     // 兜底：非法相位锁存
    _uFault := 16#0004_02AB;
    bError  := TRUE;
    _eState := E_DL_AffState.eFault;
END_CASE

(* —— 段 5｜状态出口单点映射（名实同源） —— *)
eFricZone := _eZone;
eState := _eState;
END_FUNCTION_BLOCK

(* ---- FB_DL_AxisHomeRepeatVerify.st ---- *)
(*
  Name        : FB_DL_AxisHomeRepeatVerify
  Category    : DL_Motion
  Version     : 1.0.1
  Purpose     : 回零重复性校验：收集 N 次回零到位位置，求均值/标准差/极差，散布超容差即拒绝放行（bPass = FALSE）；/ Verify homing repeatability: collect N homing positions, compute mean, standard deviation and range, and refuse release when the spread exceeds the tolerance
  溯源        : 借 t1-6-plcopen·homing 的分类/参数域组织，clean-room 实现
  Boundary    : ① 组态闸：样本数域 2..16 / 容差 <= 0 → 锁存故障（样本数 < 2 时标准差无意义）；
                ② 除子闸：标准差除子 (n-1) 恒 >= 1（n >= 2 由组态闸保证）；极差无除法；
                ③ 非有限位置该次不入样（拒收计数 bSampleRej 供诊断），不污染统计；
                ④ 完成脉冲单拍化：内部 _bDoneC 置位 → 出口统一映射（R187），不在 CASE 内直写；
                ⑤ 判定用「极差 <= 容差 且 3σ <= 容差」双条件，任一不满足即拒绝。
  修订记录    : 2026-11-20 v1.0.1：bPass/bReject 每拍预清移入 eCollect 结算拍（eDone 相保持判定，R52-02/R191）；eIdle 分支补 nGot 出口同步清零（R52-03）。
*)
TYPE E_DL_AhrState :
(
    eIdle   := 0,                            (* 未使能 / Disabled *)
    eCollect:= 10,                           (* 采样收集中 / Collecting *)
    eDone   := 20,                           (* 判定完成（等复位/等下一次启采） / Verdict done *)
    eFault  := 90                            (* 故障锁存相 / Fault latched *)
);
END_TYPE

TYPE E_DL_AhrCause :
(
    eNone       := 0,                        (* 无故障成因 / No cause *)
    eCfgIllegal := 1,                        (* 组态非法：样本数/容差越域 / Illegal config *)
    ePhaseBad   := 2                         (* 非法相位兜底 / Illegal phase fallback *)
);
END_TYPE

FUNCTION_BLOCK FB_DL_AxisHomeRepeatVerify
VAR_INPUT
    fHomePos  : REAL := 0.0;                 (* 回零到位位置（实际位置）[mm] / Homing position *)
    bHomeDone : BOOL := FALSE;               (* 单次回零完成脉冲（上升沿采一个样本）[-] / One homing done pulse *)
    nSamples  : INT := 5;                    (* 采样次数，域 2..16 [次] / Sample count, 2..16 *)
    fTolSpread: REAL := 0.05;                (* 允许散布（极差与 3σ 共用），域 > 0 [mm] / Allowed spread, > 0 *)
    bEnable   : BOOL := TRUE;                (* 校验使能 [-] / Enable *)
    bReset    : BOOL := FALSE;               (* 复位命令，上升沿清样本与判定 [-] / Reset command *)
END_VAR
VAR_OUTPUT
    nGot      : INT;                         (* 已收有效样本数 [次] / Valid samples collected *)
    fMean     : REAL;                        (* 样本均值 [mm] / Sample mean *)
    fStdDev   : REAL;                        (* 样本标准差（n-1 分母）[mm] / Sample standard deviation *)
    fSpread   : REAL;                        (* 极差 = max - min [mm] / Range *)
    bPass     : BOOL;                        (* 判定：重复性合格（可放行）[-] / Repeatability passed *)
    bReject   : BOOL;                        (* 判定：超散拒绝放行 [-] / Rejected *)
    bDone     : BOOL;                        (* 判定完成单拍脉冲 [-] / Verdict done pulse *)
    bSampleRej: BOOL;                        (* 本拍有非有限样本被拒收 [-] / Sample rejected this scan *)
    eState    : E_DL_AhrState;               (* 状态出口 / State outlet *)
    eCause    : E_DL_AhrCause;               (* 故障成因出口（R190 归因唯一） / Fault cause outlet *)
    bError    : BOOL;                        (* 故障锁存标志 [-] / Fault latch flag *)
END_VAR
VAR
    _eState  : E_DL_AhrState := E_DL_AhrState.eIdle;     (* 内部相位（CASE 唯一写入目标） / Internal phase *)
    _eCause  : E_DL_AhrCause := E_DL_AhrCause.eNone;     (* 故障成因锁存量 / Latched cause *)
    rtDone   : R_TRIG;                       (* 完成脉冲上升沿实例，段 0 无条件调用 / Homing done edge *)
    rtReset  : R_TRIG;                       (* 复位沿实例，段 0 无条件调用 / Reset edge instance *)
    _bFault  : BOOL;                         (* 故障锁存位 / Latched fault bit *)
    _bCfgBad : BOOL;                         (* 组态非法当拍量 / Illegal config this scan *)
    _bFinite : BOOL;                         (* 位置有限性当拍量 / Position finiteness *)
    _bDoneC  : BOOL;                         (* 判定完成内部单拍量（出口统一映射） / Done internal pulse *)
    _bFin    : BOOL;                         (* 本拍样本收下标志 / Sample accepted this scan *)
    _aPos    : ARRAY[1..16] OF REAL;         (* 回零位置样本数组 [mm] / Homing position samples *)
    _nGot    : INT;                          (* 样本计数 [次] / Sample counter *)
    _nIdx    : INT;                          (* 统计游标（每趟重置，R227）[-] / Stats cursor *)
    _nEff    : INT;                          (* 钳位后生效样本数 [次] / Clamped sample count *)
    _fSum    : REAL;                         (* Σx [mm] / Sum *)
    _fMeanI  : REAL;                         (* 均值中间量 [mm] / Mean intermediate *)
    _fVar    : REAL;                         (* Σ(x-x̄)² [mm²] / Sum of squares *)
    _fMin    : REAL;                         (* 样本最小值 [mm] / Minimum *)
    _fMax    : REAL;                         (* 样本最大值 [mm] / Maximum *)
    _fStd    : REAL;                         (* 标准差中间量 [mm] / Std intermediate *)
END_VAR
VAR CONSTANT
    DL_AHR_EPS   : REAL := 1.0E-6;           (* 判零容差 [-] / Epsilon *)
    DL_AHR_NMAX  : INT  := 16;               (* 样本容量上限 [次] / Sample capacity *)
    DL_AHR_NMIN  : INT  := 2;                (* 样本数下限（标准差最少两点）[次] / Sample lower bound *)
    DL_AHR_SIGMA : REAL := 3.0;              (* 散布判据 σ 倍数（3σ 工程惯例）[-] / Sigma multiplier *)
END_VAR

(* —— 段 0：当拍判据派生 + 实例无条件刷新（R228A） —— *)
_bCfgBad := (nSamples < DL_AHR_NMIN) OR (nSamples > DL_AHR_NMAX)               (* 样本数域闸 / Sample-count gate *)
            OR (fTolSpread <= DL_AHR_EPS);                                     (* 容差正域闸 / Tolerance gate *)
rtDone(CLK := bHomeDone);                                                      (* 完成沿每拍必调 / Done edge every scan *)
rtReset(CLK := bReset);                                                        (* 复位沿每拍必调 / Reset edge every scan *)
_bFinite := (fHomePos = fHomePos) AND ((fHomePos - fHomePos) = (fHomePos - fHomePos));   (* NaN 自反 + Inf 差判 / NaN and Inf gate *)
_nEff := nSamples;                                                             (* 生效样本数初值 / Effective count *)
IF _nEff < DL_AHR_NMIN THEN
    _nEff := DL_AHR_NMIN;                                                      (* 下限钳位 / Lower clamp *)
END_IF
IF _nEff > DL_AHR_NMAX THEN
    _nEff := DL_AHR_NMAX;                                                      (* 上限钳位（R308） / Upper clamp *)
END_IF

(* —— 段 1：单拍量预清零（R107） —— *)
_bDoneC := FALSE;                                                              (* 完成脉冲内部量预清 / Done preset *)
bSampleRej := FALSE;                                                           (* 拒收指示预清 / Reject-sample preset *)

(* —— 段 2：复位沿处理（作用域：清故障 + 清样本 + 清统计 + 迁 eIdle，R283 逐项声明） —— *)
IF rtReset.Q THEN
    _bFault := FALSE;                                                          (* 清故障锁存 / Clear fault *)
    _eCause := E_DL_AhrCause.eNone;                                            (* 清成因 / Clear cause *)
    _nGot := 0;                                                                (* 清样本计数 / Clear sample counter *)
    nGot := 0;                                                                 (* 清出口计数 / Clear outlet count *)
    fMean := 0.0;                                                              (* 清均值出口 / Clear mean *)
    fStdDev := 0.0;                                                            (* 清标准差出口 / Clear std *)
    fSpread := 0.0;                                                            (* 清极差出口 / Clear range *)
    _eState := E_DL_AhrState.eIdle;                                            (* 迁未使能相 / Back to idle *)
END_IF

(* —— 段 3：组态故障锁存（锁存至复位沿，R189） —— *)
IF _bCfgBad AND NOT _bFault THEN
    _bFault := TRUE;                                                           (* 锁存故障位 / Latch fault *)
    _eCause := E_DL_AhrCause.eCfgIllegal;                                      (* 成因：组态非法 / Cause: illegal config *)
    _eState := E_DL_AhrState.eFault;                                           (* 同步迁故障相 / Migrate to fault *)
END_IF

(* —— 段 4：CASE 主状态机（ELSE 兜底迁 eFault，红线 6） —— *)
CASE _eState OF
    E_DL_AhrState.eIdle:                                                       (* 未使能：不采样 / Disabled *)
        _nGot := 0;                                                            (* 失能清样本计数（防隐性回夹） / Clear sample counter *)
        nGot := 0;                                                             (* 失能同步清出口计数（R52-03 名实一致） / Clear outlet count *)
        bPass := FALSE;                                                        (* 失能清判定出口（复位/失能路径出口清零） / Clear verdict outlets *)
        bReject := FALSE;                                                      (* 失能清拒绝出口 / Clear reject outlet *)
        IF bEnable AND NOT _bFault THEN
            _eState := E_DL_AhrState.eCollect;                                 (* 使能进入收集 / Enter collecting *)
        END_IF
    E_DL_AhrState.eCollect:                                                    (* 收集相：逐次入样 / Collecting *)
        IF NOT bEnable THEN
            _eState := E_DL_AhrState.eIdle;                                    (* 失能回未使能 / Back to idle *)
        ELSIF rtDone.Q THEN                                                    (* 一次回零完成 / One homing done *)
            _bFin := _bFinite;                                                 (* 本拍样本有效性 / Sample validity *)
            IF _bFin AND (_nGot < DL_AHR_NMAX) THEN
                _nGot := _nGot + 1;                                            (* 计数先增（<= 容量闸） / Count up within capacity *)
                _aPos[_nGot] := fHomePos;                                      (* 入样（下标已由容量闸限住） / Store sample *)
                nGot := _nGot;                                                 (* 出口计数镜像 / Outlet mirror *)
            ELSIF NOT _bFin THEN
                bSampleRej := TRUE;                                            (* 非有限样本拒收（边界③） / Reject non-finite *)
            END_IF
        END_IF
        IF _nGot >= _nEff THEN                                                 (* 样本到齐：一次性统计 / Enough samples: compute *)
            _fSum := 0.0;                                                      (* Σx 预清 / Sum preset *)
            _nIdx := 1;                                                        (* 游标起头（R227） / Cursor reset *)
            _fMin := _aPos[1];                                                 (* 最小值初值取首样本 / Min init *)
            _fMax := _aPos[1];                                                 (* 最大值初值取首样本 / Max init *)
            WHILE _nIdx <= _nEff DO                                            (* 一趟求 Σx/min/max（下标已钳位） / One pass for sum/min/max *)
                _fSum := _fSum + _aPos[_nIdx];                                 (* Σx [mm] / Sum *)
                IF _aPos[_nIdx] < _fMin THEN
                    _fMin := _aPos[_nIdx];                                     (* 更新最小值 / Update min *)
                END_IF
                IF _aPos[_nIdx] > _fMax THEN
                    _fMax := _aPos[_nIdx];                                     (* 更新最大值 / Update max *)
                END_IF
                _nIdx := _nIdx + 1;                                            (* 游标递进 / Cursor advance *)
            END_WHILE
            _fMeanI := _fSum / DINT_TO_REAL(_nEff);                            (* 均值：除子 nEff >= 2 无除零 [mm] / Mean, divisor >= 2 *)
            fMean := _fMeanI;                                                  (* 均值出口 / Mean outlet *)
            fSpread := _fMax - _fMin;                                          (* 极差（无除法）[mm] / Range *)
            _fVar := 0.0;                                                      (* 平方和预清 / Squares preset *)
            _nIdx := 1;                                                        (* 游标重起 / Cursor reset *)
            WHILE _nIdx <= _nEff DO                                            (* 二趟求 Σ(x-x̄)² / Second pass for variance *)
                _fVar := _fVar + (_aPos[_nIdx] - _fMeanI) * (_aPos[_nIdx] - _fMeanI);   (* 平方项恒非负 [mm²] / Squared deviation *)
                _nIdx := _nIdx + 1;                                            (* 游标递进 / Cursor advance *)
            END_WHILE
            _fStd := SQRT(_fVar / DINT_TO_REAL(_nEff - 1));                    (* 样本标准差：除子 nEff-1 >= 1 [mm] / Sample std, divisor >= 1 *)
            fStdDev := _fStd;                                                  (* 标准差出口 / Std outlet *)
            bPass := FALSE;                                                    (* 结算拍预清合格位（当拍二选一赋值，eDone 相保持） / Preset pass at settle scan *)
            bReject := FALSE;                                                  (* 结算拍预清拒绝位 / Preset reject at settle scan *)
            IF (fSpread <= fTolSpread) AND ((DL_AHR_SIGMA * _fStd) <= fTolSpread) THEN
                bPass := TRUE;                                                 (* 双条件满足：重复性合格 / Both conditions met: pass *)
            ELSE
                bReject := TRUE;                                               (* 任一不满足：超散拒绝放行 / Reject on spread *)
            END_IF
            _bDoneC := TRUE;                                                   (* 完成脉冲内部置位（出口统一映射，R187） / Done pulse internal *)
            _eState := E_DL_AhrState.eDone;                                    (* 迁完成相 / To done *)
        END_IF
    E_DL_AhrState.eDone:                                                       (* 完成相：保持判定，等复位或重新使能 / Done *)
        IF NOT bEnable THEN
            _eState := E_DL_AhrState.eIdle;                                    (* 失能回未使能 / Back to idle *)
        END_IF
    E_DL_AhrState.eFault:                                                      (* 故障相：冻结保持末值，仅复位沿出 / Fault *)
        ;                                                                      (* 锁存回放（R28） / Replay from latch *)
    ELSE                                                                       (* 非法相位兜底迁安全态 / Illegal phase fallback *)
        _eState := E_DL_AhrState.eFault;                                       (* 迁故障相 / To fault *)
        _bFault := TRUE;                                                       (* 同步锁存 / Latch *)
        _eCause := E_DL_AhrCause.ePhaseBad;                                    (* 成因：非法相位 / Cause: illegal phase *)
END_CASE

(* —— 段 5：出口映射（内部 _b* → 输出单拍，R187；名实双出口，R191） —— *)
bDone := _bDoneC;                                                              (* 完成脉冲单拍出口 / Done single-scan outlet *)
bError := _bFault;                                                             (* 故障标志镜像 / Fault flag mirror *)
eState := _eState;                                                             (* 状态出口 / State outlet *)
eCause := _eCause;                                                             (* 成因出口 / Cause outlet *)
END_FUNCTION_BLOCK
